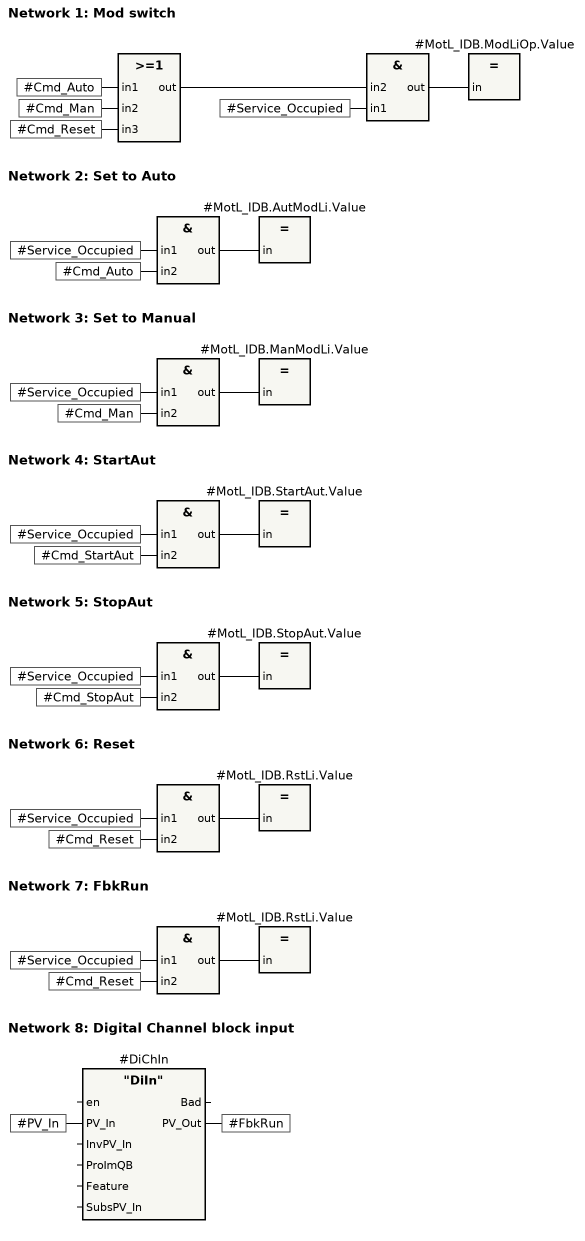
   #MotL_IDB.ModLiOp.Value := (#Cmd_Auto OR #Cmd_Man OR #Cmd_Reset) AND #Service_Occupied;
END_REGION

REGION Network 2: Set to Auto
   #MotL_IDB.AutModLi.Value := #Service_Occupied AND #Cmd_Auto;
END_REGION

REGION Network 3: Set to Manual
   #MotL_IDB.ManModLi.Value := #Service_Occupied AND #Cmd_Man;
END_REGION

REGION Network 4: StartAut
   #MotL_IDB.StartAut.Value := #Service_Occupied AND #Cmd_StartAut;
END_REGION

REGION Network 5: StopAut
   #MotL_IDB.StopAut.Value := #Service_Occupied AND #Cmd_StopAut;
END_REGION

REGION Network 6: Reset
   #MotL_IDB.RstLi.Value := #Service_Occupied AND #Cmd_Reset;
END_REGION

REGION Network 7: FbkRun
   #MotL_IDB.RstLi.Value := #Service_Occupied AND #Cmd_Reset;
END_REGION

REGION Network 8: Digital Channel block input
   #DiChIn(PV_In := #PV_In, PV_Out => #FbkRun);   // "DiIn"
END_REGION

REGION Network 9: CSF
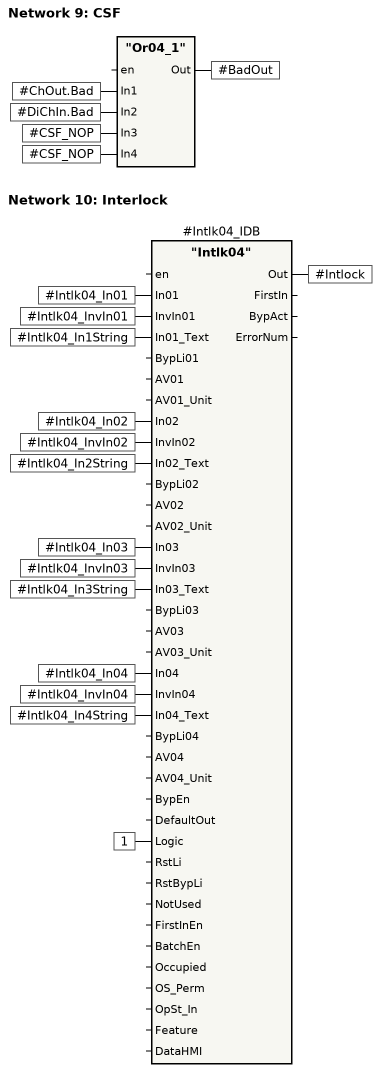
   "Or04_1"(In1 := #ChOut.Bad, In2 := #DiChIn.Bad, In3 := #CSF_NOP, In4 := #CSF_NOP, Out => #BadOut);
END_REGION

REGION Network 10: Interlock
   #Intlk04_IDB(In01 := #Intlk04_In01,   // "Intlk04"
                InvIn01 := #Intlk04_InvIn01,
                In01_Text := #Intlk04_In1String,
                In02 := #Intlk04_In02,
                InvIn02 := #Intlk04_InvIn02,
                In02_Text := #Intlk04_In2String,
                In03 := #Intlk04_In03,
                InvIn03 := #Intlk04_InvIn03,
                In03_Text := #Intlk04_In3String,
                In04 := #Intlk04_In04,
                InvIn04 := #Intlk04_InvIn04,
                In04_Text := #Intlk04_In4String,
                Logic := 1,
                Out => #Intlock);
END_REGION

REGION Network 11: MotSpdCL
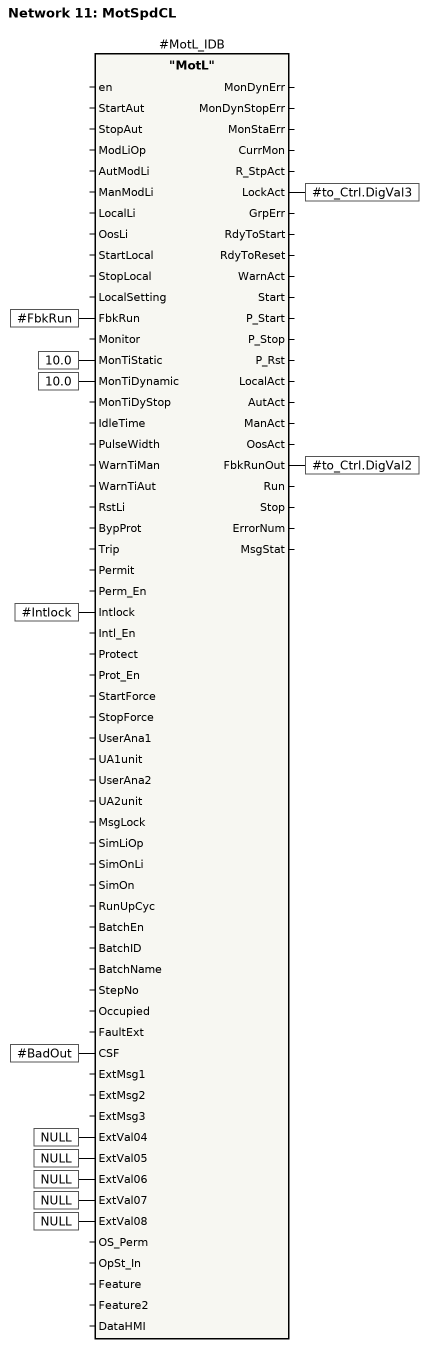
   #MotL_IDB(FbkRun := #FbkRun,   // "MotL"
             MonTiStatic := 10.0,
             MonTiDynamic := 10.0,
             Intlock := #Intlock,
             CSF := #BadOut,
             ExtVal04 := NULL,
             ExtVal05 := NULL,
             ExtVal06 := NULL,
             ExtVal07 := NULL,
             ExtVal08 := NULL,
             LockAct => #to_Ctrl.DigVal3,
             FbkRunOut => #to_Ctrl.DigVal2);
END_REGION

REGION Network 12: Channel block output
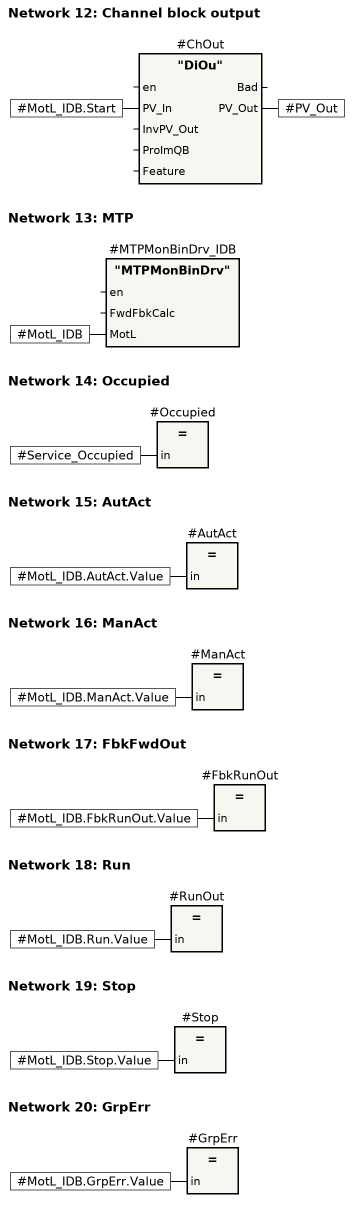
   #ChOut(PV_In := #MotL_IDB.Start, PV_Out => #PV_Out);   // "DiOu"
END_REGION

REGION Network 13: MTP
   #MTPMonBinDrv_IDB(MotL := #MotL_IDB);   // "MTPMonBinDrv"
END_REGION

REGION Network 14: Occupied
   #Occupied := #Service_Occupied;
END_REGION

REGION Network 15: AutAct
   #AutAct := #MotL_IDB.AutAct.Value;
END_REGION

REGION Network 16: ManAct
   #ManAct := #MotL_IDB.ManAct.Value;
END_REGION

REGION Network 17: FbkFwdOut
   #FbkRunOut := #MotL_IDB.FbkRunOut.Value;
END_REGION

REGION Network 18: Run
   #RunOut := #MotL_IDB.Run.Value;
END_REGION

REGION Network 19: Stop
   #Stop := #MotL_IDB.Stop.Value;
END_REGION

REGION Network 20: GrpErr
   #GrpErr := #MotL_IDB.GrpErr.Value;
END_REGION
END_FUNCTION_BLOCK

FUNCTION "P101" : Void   // FC17, FBD
{ S7_Optimized_Access := 'TRUE' }
// stored: SetENOAutomatically false
   VAR_TEMP
      Temp : "DigVal";
      Temp_1 : "DigVal";
      Temp_3 : "DigVal";
      Temp_2 : "DigVal";
      Temp_Error : "DigVal";
      In03 : "DigVal";
      State : "Service_States";
      FbkRun : "DigVal";
      StopAut : Bool;
   END_VAR
   VAR_TEMP   // added for the SCL form of the ladder/FBD networks
      _w1 : Bool;
   END_VAR
BEGIN

REGION Network 1: simulate Fbk Error
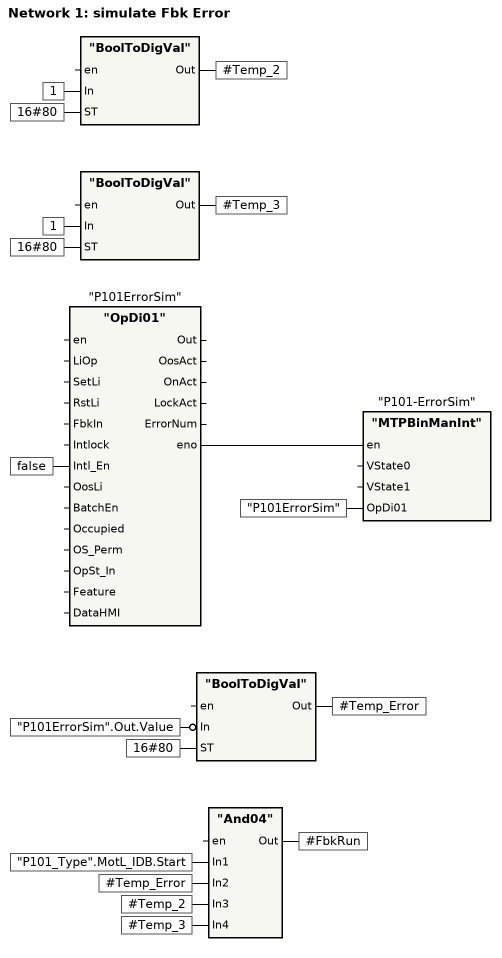
   "BoolToDigVal"(In := 1, ST := 16#80, Out => #Temp_2);
   "BoolToDigVal"(In := 1, ST := 16#80, Out => #Temp_3);
   "P101ErrorSim"(Intl_En := false, ENO => #_w1);   // "OpDi01"
   IF #_w1 THEN
       "P101-ErrorSim"(OpDi01 := "P101ErrorSim");   // "MTPBinManInt"
   END_IF;
   "BoolToDigVal"(In := NOT "P101ErrorSim".Out.Value, ST := 16#80, Out => #Temp_Error);
   "And04"(In1 := "P101_Type".MotL_IDB.Start,
           In2 := #Temp_Error,
           In3 := #Temp_2,
           In4 := #Temp_3,
           Out => #FbkRun);
END_REGION

REGION Network 2: Pump interconnections
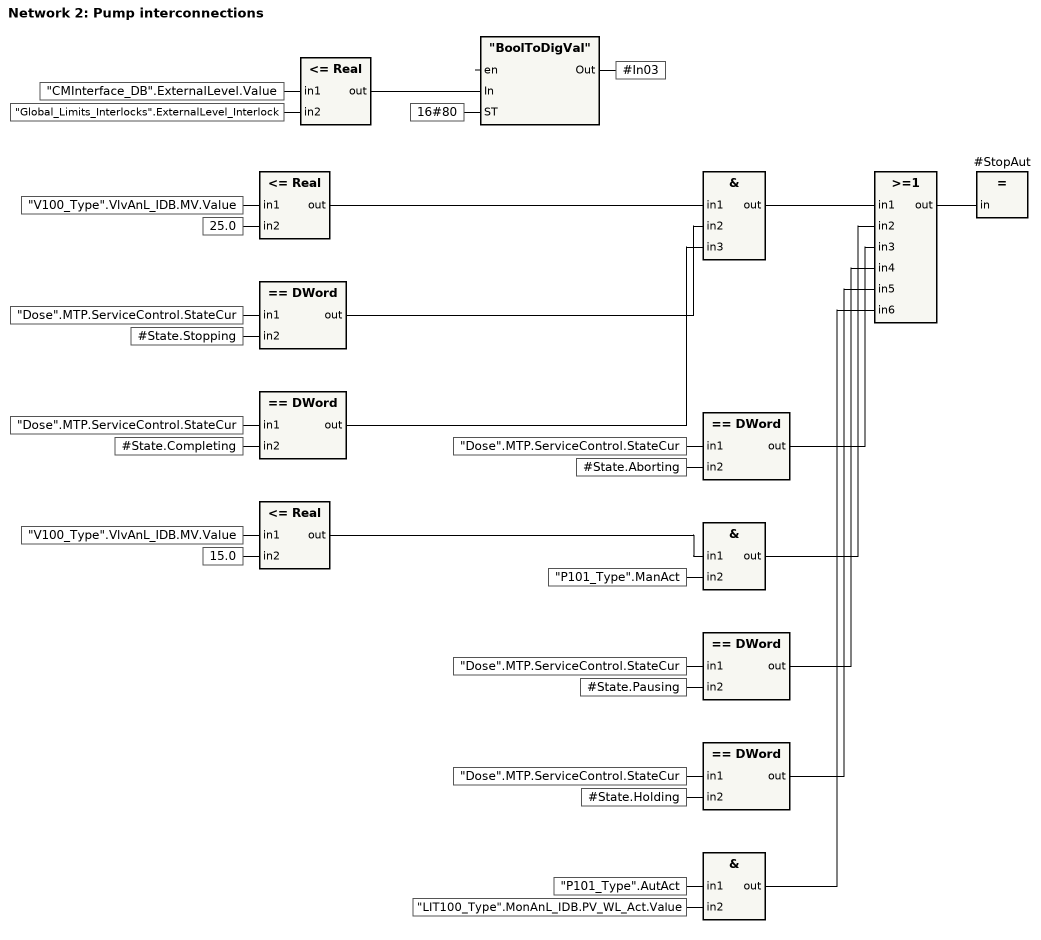
   "BoolToDigVal"(In := "CMInterface_DB".ExternalLevel.Value <= "Global_Limits_Interlocks".ExternalLevel_Interlock,
                  ST := 16#80,
                  Out => #In03);
   #StopAut := (("V100_Type".VlvAnL_IDB.MV.Value <= 25.0) AND ("Dose".MTP.ServiceControl.StateCur = #State.Stopping) AND ("Dose".MTP.ServiceControl.StateCur = #State.Completing)) OR (("V100_Type".VlvAnL_IDB.MV.Value <= 15.0) AND "P101_Type".ManAct) OR ("Dose".MTP.ServiceControl.StateCur = #State.Aborting) OR ("Dose".MTP.ServiceControl.StateCur = #State.Pausing) OR ("Dose".MTP.ServiceControl.StateCur = #State.Holding) OR ("P101_Type".AutAct AND "LIT100_Type".MonAnL_IDB.PV_WL_Act.Value);
END_REGION

REGION Network 3: MotL
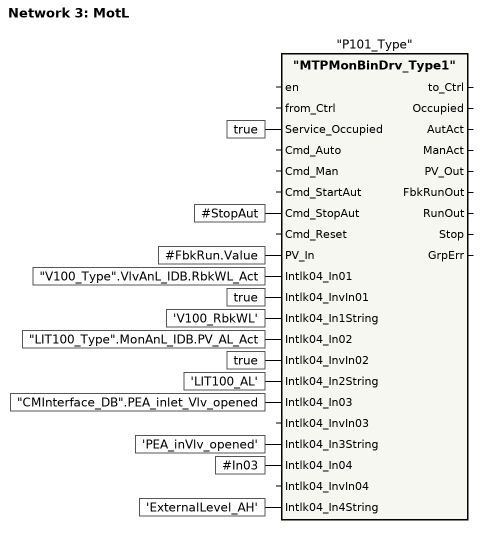
   "P101_Type"(Service_Occupied := true,   // "MTPMonBinDrv_Type1"
               Cmd_StopAut := #StopAut,
               PV_In := #FbkRun.Value,
               Intlk04_In01 := "V100_Type".VlvAnL_IDB.RbkWL_Act,
               Intlk04_InvIn01 := true,
               Intlk04_In1String := 'V100_RbkWL',
               Intlk04_In02 := "LIT100_Type".MonAnL_IDB.PV_AL_Act,
               Intlk04_InvIn02 := true,
               Intlk04_In2String := 'LIT100_AL',
               Intlk04_In03 := "CMInterface_DB".PEA_inlet_Vlv_opened,
               Intlk04_In3String := 'PEA_inVlv_opened',
               Intlk04_In04 := #In03,
               Intlk04_In4String := 'ExternalLevel_AH');
END_REGION
END_FUNCTION

FUNCTION "V100" : Void   // FC3, FBD
{ S7_Optimized_Access := 'TRUE' }
// stored: SetENOAutomatically false
   VAR_TEMP
      Temp : "DigVal";
      In03 : "DigVal";
      Temp_FF : "DigVal";
      Temp_fromCTRL : "StruCm";
   END_VAR
BEGIN

REGION Network 1: VlvAnL interconnections
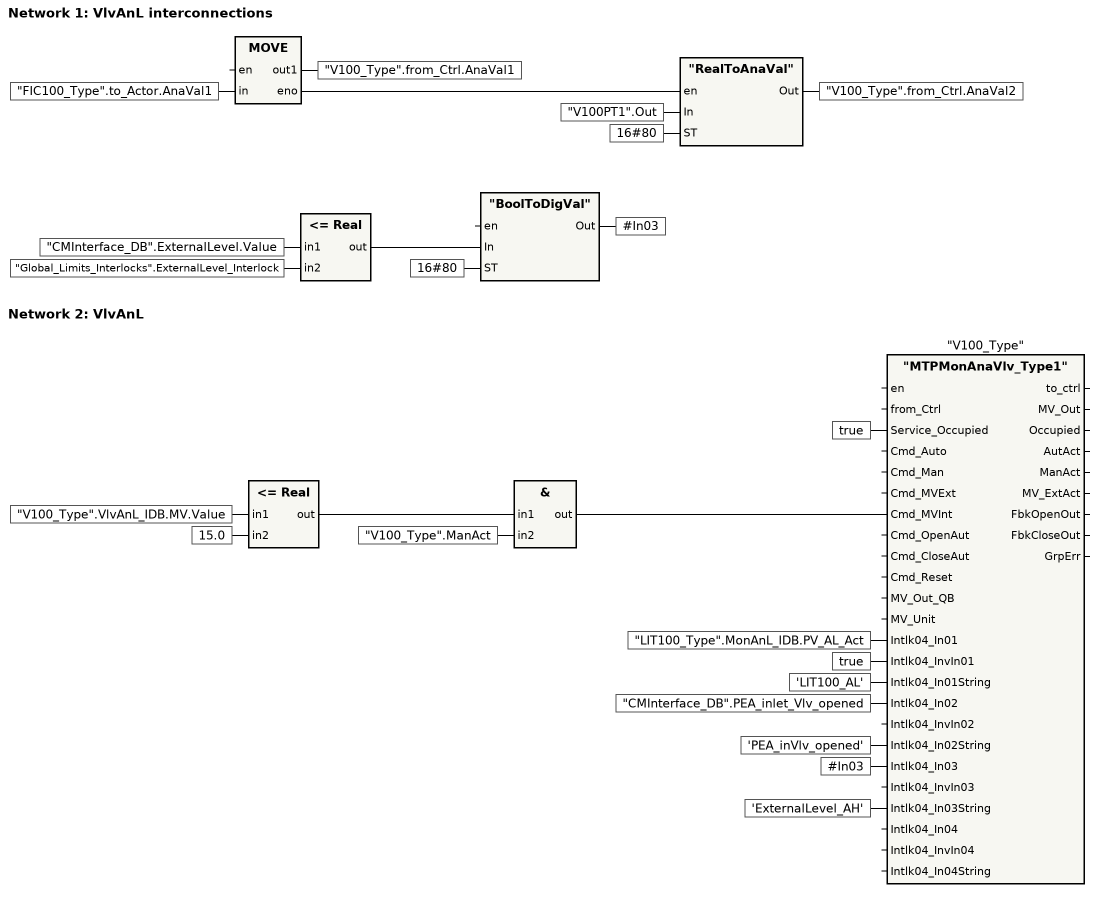
   "V100_Type".from_Ctrl.AnaVal1 := "FIC100_Type".to_Actor.AnaVal1;
   "RealToAnaVal"(In := "V100PT1".Out, ST := 16#80, Out => "V100_Type".from_Ctrl.AnaVal2);
   "BoolToDigVal"(In := "CMInterface_DB".ExternalLevel.Value <= "Global_Limits_Interlocks".ExternalLevel_Interlock,
                  ST := 16#80,
                  Out => #In03);
END_REGION

REGION Network 2: VlvAnL
   "V100_Type"(Service_Occupied := true,   // "MTPMonAnaVlv_Type1"
               Cmd_MVInt := ("V100_Type".VlvAnL_IDB.MV.Value <= 15.0) AND "V100_Type".ManAct,
               Intlk04_In01 := "LIT100_Type".MonAnL_IDB.PV_AL_Act,
               Intlk04_InvIn01 := true,
               Intlk04_In01String := 'LIT100_AL',
               Intlk04_In02 := "CMInterface_DB".PEA_inlet_Vlv_opened,
               Intlk04_In02String := 'PEA_inVlv_opened',
               Intlk04_In03 := #In03,
               Intlk04_In03String := 'ExternalLevel_AH');
END_REGION
END_FUNCTION

FUNCTION "RealToAnaVal" : Void   // FC9, SCL
{ S7_Optimized_Access := 'TRUE' }
// stored: SetENOAutomatically false
   VAR_INPUT
      In : Real;
      ST : Byte;
   END_VAR
   VAR_OUTPUT
      Out : "AnaVal";
   END_VAR
BEGIN
   #Out.ST := #ST;
   #Out.Value := #In;
END_FUNCTION

FUNCTION_BLOCK "MTPMonAnaVlv_Type1"   // FB7, FBD
{ S7_Optimized_Access := 'TRUE' }
// stored: MemoryReserve 100, SetENOAutomatically false
   VAR_INPUT
      from_Ctrl { ExternalAccessible := 'False'; ExternalVisible := 'False'; ExternalWritable := 'False'} : "StruCm";
      Service_Occupied { ExternalAccessible := 'False'; ExternalVisible := 'False'; ExternalWritable := 'False'} : Bool;
      Cmd_Auto { ExternalAccessible := 'False'; ExternalVisible := 'False'; ExternalWritable := 'False'} : Bool;
      Cmd_Man { ExternalAccessible := 'False'; ExternalVisible := 'False'; ExternalWritable := 'False'} : Bool;
      Cmd_MVExt { ExternalAccessible := 'False'; ExternalVisible := 'False'; ExternalWritable := 'False'} : Bool;
      Cmd_MVInt { ExternalAccessible := 'False'; ExternalVisible := 'False'; ExternalWritable := 'False'} : Bool;
      Cmd_OpenAut { ExternalAccessible := 'False'; ExternalVisible := 'False'; ExternalWritable := 'False'} : Bool;
      Cmd_CloseAut { ExternalAccessible := 'False'; ExternalVisible := 'False'; ExternalWritable := 'False'} : Bool;
      Cmd_Reset { ExternalAccessible := 'False'; ExternalVisible := 'False'; ExternalWritable := 'False'} : Bool;
      MV_Out_QB { ExternalAccessible := 'False'; ExternalVisible := 'False'; ExternalWritable := 'False'} : Bool := true;
      MV_Unit { ExternalAccessible := 'False'; ExternalVisible := 'False'; ExternalWritable := 'False'} : Int := 1342;
      Intlk04_In01 { ExternalAccessible := 'False'; ExternalVisible := 'False'; ExternalWritable := 'False'} : "DigVal";
      Intlk04_InvIn01 { ExternalAccessible := 'False'; ExternalVisible := 'False'; ExternalWritable := 'False'} : Bool;
      Intlk04_In01String : String;
      Intlk04_In02 { ExternalAccessible := 'False'; ExternalVisible := 'False'; ExternalWritable := 'False'} : "DigVal";
      Intlk04_InvIn02 { ExternalAccessible := 'False'; ExternalVisible := 'False'; ExternalWritable := 'False'} : Bool;
      Intlk04_In02String : String;
      Intlk04_In03 { ExternalAccessible := 'False'; ExternalVisible := 'False'; ExternalWritable := 'False'} : "DigVal";
      Intlk04_InvIn03 { ExternalAccessible := 'False'; ExternalVisible := 'False'; ExternalWritable := 'False'} : Bool;
      Intlk04_In03String : String;
      Intlk04_In04 { ExternalAccessible := 'False'; ExternalVisible := 'False'; ExternalWritable := 'False'} : "DigVal";
      Intlk04_InvIn04 { ExternalAccessible := 'False'; ExternalVisible := 'False'; ExternalWritable := 'False'} : Bool;
      Intlk04_In04String : String;
   END_VAR
   VAR_OUTPUT
      to_ctrl { ExternalAccessible := 'False'; ExternalVisible := 'False'; ExternalWritable := 'False'} : "StruCm";
      MV_Out { ExternalAccessible := 'False'; ExternalVisible := 'False'; ExternalWritable := 'False'} : Word;
      Occupied { ExternalAccessible := 'False'; ExternalVisible := 'False'; ExternalWritable := 'False'} : Bool;   // Occupied by a Service procedure
      AutAct { ExternalAccessible := 'False'; ExternalVisible := 'False'; ExternalWritable := 'False'} : Bool;
      ManAct { ExternalAccessible := 'False'; ExternalVisible := 'False'; ExternalWritable := 'False'} : Bool;
      MV_ExtAct { ExternalAccessible := 'False'; ExternalVisible := 'False'; ExternalWritable := 'False'} : Bool;
      FbkOpenOut { ExternalAccessible := 'False'; ExternalVisible := 'False'; ExternalWritable := 'False'} : Bool;
      FbkCloseOut { ExternalAccessible := 'False'; ExternalVisible := 'False'; ExternalWritable := 'False'} : Bool;
      GrpErr { ExternalAccessible := 'False'; ExternalVisible := 'False'; ExternalWritable := 'False'} : Bool;
   END_VAR
   VAR
      AnOut_IDB { ExternalAccessible := 'False'; ExternalVisible := 'False'; ExternalWritable := 'False'} : "AnOu";
      Intlk04_IDB : "Intlk04";
      VlvAnL_IDB { S7_SetPoint := 'True'} : "VlvAnL";
      MTPMonAnaVlv_IDB { ExternalVisible := 'False'; S7_SetPoint := 'True'} : "MTPMonAnaVlv";
   END_VAR
   VAR_TEMP
      CSF_NOP : "DigVal";
      BadAnIn : "DigVal";
      BadOut : "DigVal";
      Intlock : "DigVal";
   END_VAR
   // Intlk04_In01.Value := true;
   // Intlk04_In02.Value := true;
   // Intlk04_In03.Value := true;
   // Intlk04_In04.Value := true;
BEGIN

REGION Network 1: Convert
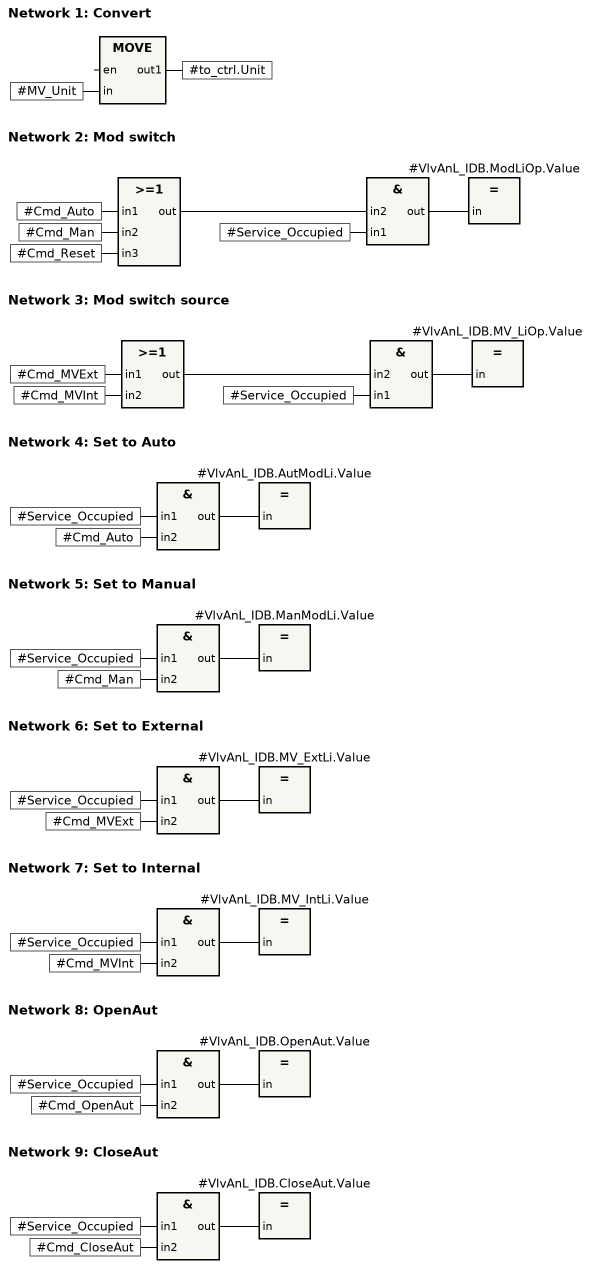
   #to_ctrl.Unit := #MV_Unit;
END_REGION

REGION Network 2: Mod switch
   #VlvAnL_IDB.ModLiOp.Value := (#Cmd_Auto OR #Cmd_Man OR #Cmd_Reset) AND #Service_Occupied;
END_REGION

REGION Network 3: Mod switch source
   #VlvAnL_IDB.MV_LiOp.Value := (#Cmd_MVExt OR #Cmd_MVInt) AND #Service_Occupied;
END_REGION

REGION Network 4: Set to Auto
   #VlvAnL_IDB.AutModLi.Value := #Service_Occupied AND #Cmd_Auto;
END_REGION

REGION Network 5: Set to Manual
   #VlvAnL_IDB.ManModLi.Value := #Service_Occupied AND #Cmd_Man;
END_REGION

REGION Network 6: Set to External
   #VlvAnL_IDB.MV_ExtLi.Value := #Service_Occupied AND #Cmd_MVExt;
END_REGION

REGION Network 7: Set to Internal
   #VlvAnL_IDB.MV_IntLi.Value := #Service_Occupied AND #Cmd_MVInt;
END_REGION

REGION Network 8: OpenAut
   #VlvAnL_IDB.OpenAut.Value := #Service_Occupied AND #Cmd_OpenAut;
END_REGION

REGION Network 9: CloseAut
   #VlvAnL_IDB.CloseAut.Value := #Service_Occupied AND #Cmd_CloseAut;
END_REGION

REGION Network 10: Reset
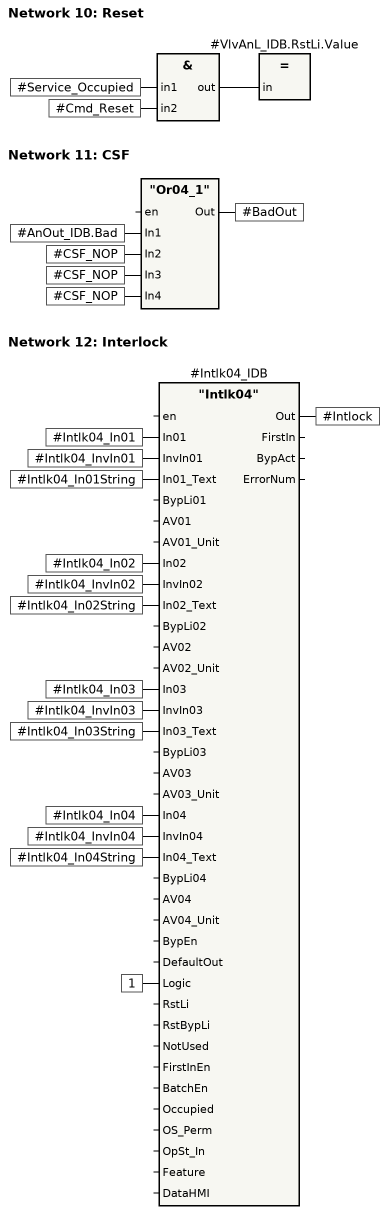
   #VlvAnL_IDB.RstLi.Value := #Service_Occupied AND #Cmd_Reset;
END_REGION

REGION Network 11: CSF
   "Or04_1"(In1 := #AnOut_IDB.Bad, In2 := #CSF_NOP, In3 := #CSF_NOP, In4 := #CSF_NOP, Out => #BadOut);
END_REGION

REGION Network 12: Interlock
   #Intlk04_IDB(In01 := #Intlk04_In01,   // "Intlk04"
                InvIn01 := #Intlk04_InvIn01,
                In01_Text := #Intlk04_In01String,
                In02 := #Intlk04_In02,
                InvIn02 := #Intlk04_InvIn02,
                In02_Text := #Intlk04_In02String,
                In03 := #Intlk04_In03,
                InvIn03 := #Intlk04_InvIn03,
                In03_Text := #Intlk04_In03String,
                In04 := #Intlk04_In04,
                InvIn04 := #Intlk04_InvIn04,
                In04_Text := #Intlk04_In04String,
                Logic := 1,
                Out => #Intlock);
END_REGION

REGION Network 13: VlvAnL
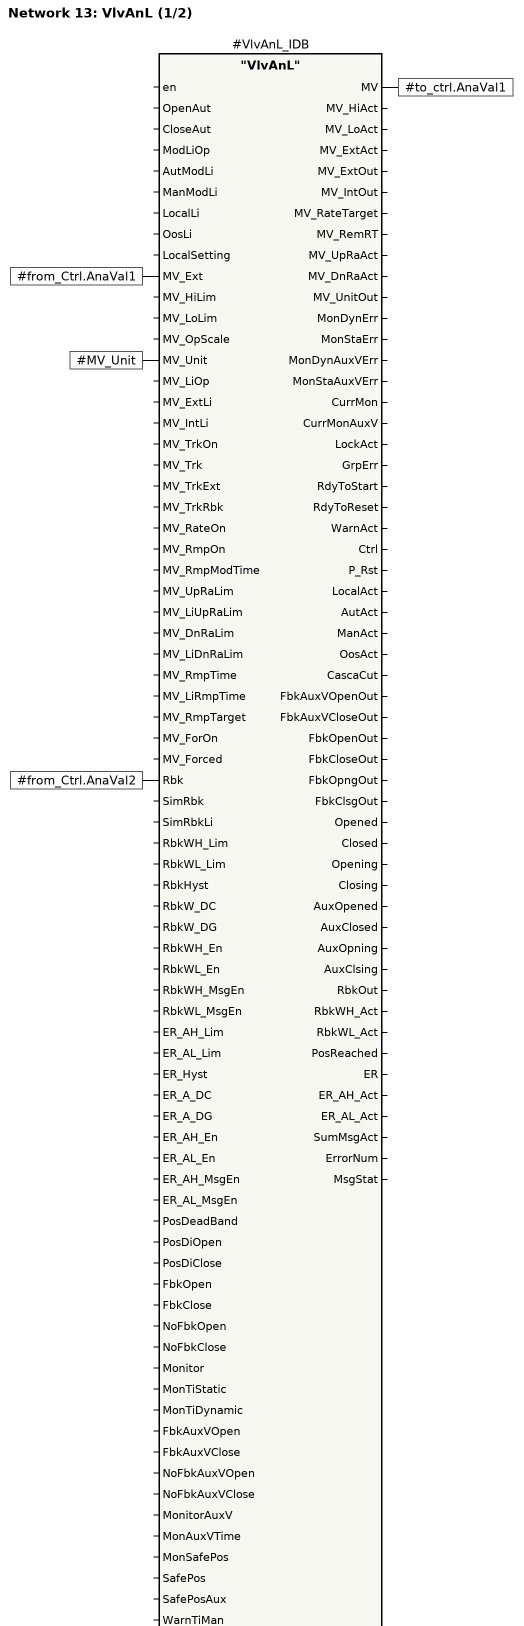
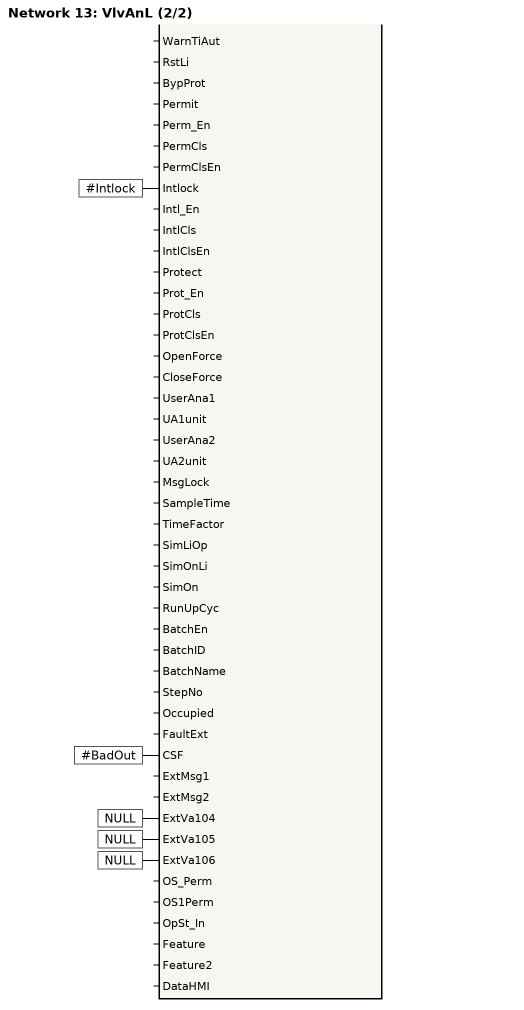
   #VlvAnL_IDB(MV_Ext := #from_Ctrl.AnaVal1,   // "VlvAnL"
               MV_Unit := #MV_Unit,
               Rbk := #from_Ctrl.AnaVal2,
               Intlock := #Intlock,
               CSF := #BadOut,
               ExtVa104 := NULL,
               ExtVa105 := NULL,
               ExtVa106 := NULL,
               MV => #to_ctrl.AnaVal1);
END_REGION

REGION Network 14: Analog Out
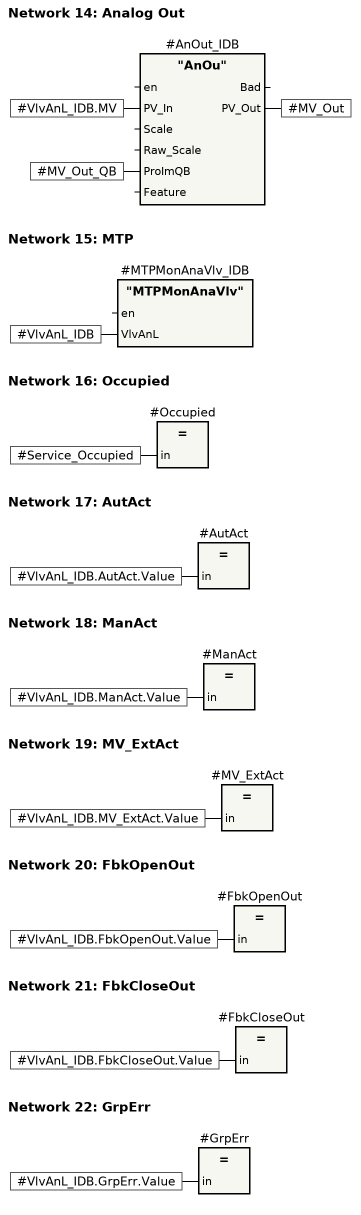
   #AnOut_IDB(PV_In := #VlvAnL_IDB.MV, ProImQB := #MV_Out_QB, PV_Out => #MV_Out);   // "AnOu"
END_REGION

REGION Network 15: MTP
   #MTPMonAnaVlv_IDB(VlvAnL := #VlvAnL_IDB);   // "MTPMonAnaVlv"
END_REGION

REGION Network 16: Occupied
   #Occupied := #Service_Occupied;
END_REGION

REGION Network 17: AutAct
   #AutAct := #VlvAnL_IDB.AutAct.Value;
END_REGION

REGION Network 18: ManAct
   #ManAct := #VlvAnL_IDB.ManAct.Value;
END_REGION

REGION Network 19: MV_ExtAct
   #MV_ExtAct := #VlvAnL_IDB.MV_ExtAct.Value;
END_REGION

REGION Network 20: FbkOpenOut
   #FbkOpenOut := #VlvAnL_IDB.FbkOpenOut.Value;
END_REGION

REGION Network 21: FbkCloseOut
   #FbkCloseOut := #VlvAnL_IDB.FbkCloseOut.Value;
END_REGION

REGION Network 22: GrpErr
   #GrpErr := #VlvAnL_IDB.GrpErr.Value;
END_REGION
END_FUNCTION_BLOCK

FUNCTION "Flow_Sim" : Void   // FC14, FBD
{ S7_Optimized_Access := 'TRUE' }
// stored: SetENOAutomatically false
   VAR_TEMP
      State : "Service_States";
   END_VAR
BEGIN

REGION Network 1: flow value
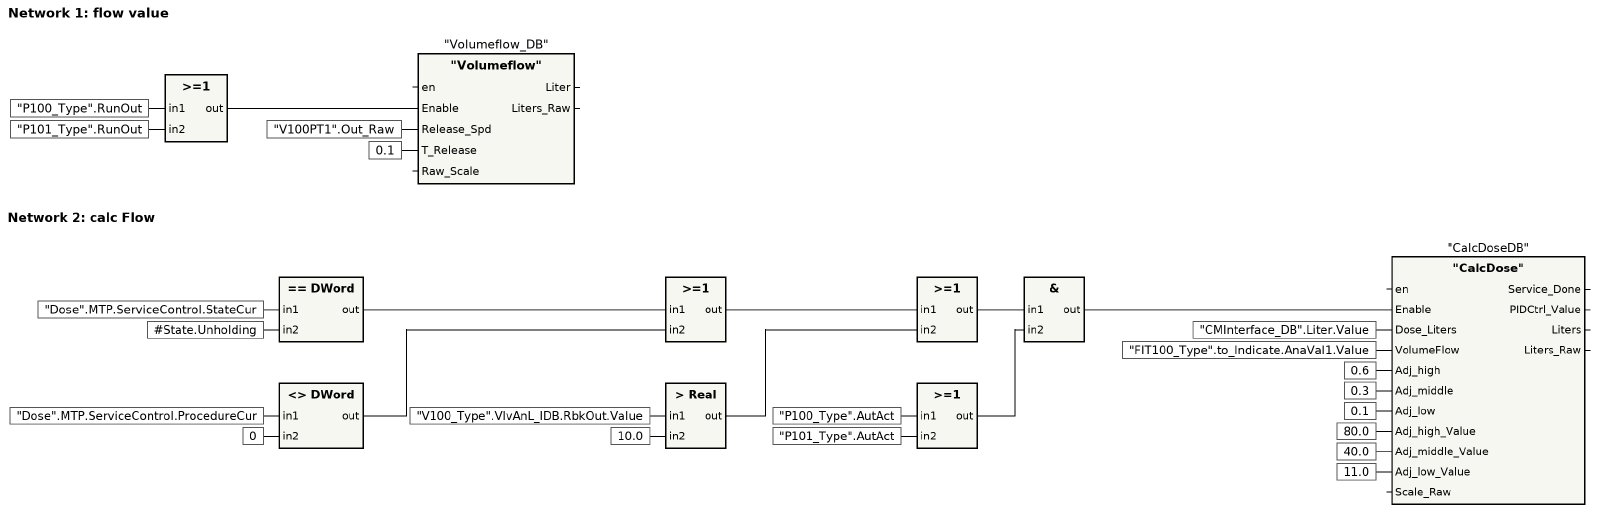
   "Volumeflow_DB"(Enable := "P100_Type".RunOut OR "P101_Type".RunOut,   // "Volumeflow"
                   Release_Spd := "V100PT1".Out_Raw,
                   T_Release := 0.1);
END_REGION

REGION Network 2: calc Flow
   "CalcDoseDB"(Enable := (("Dose".MTP.ServiceControl.StateCur = #State.Unholding) OR ("Dose".MTP.ServiceControl.ProcedureCur <> 0) OR ("V100_Type".VlvAnL_IDB.RbkOut.Value > 10.0)) AND ("P100_Type".AutAct OR "P101_Type".AutAct),   // "CalcDose"
                Dose_Liters := "CMInterface_DB".Liter.Value,
                VolumeFlow := "FIT100_Type".to_Indicate.AnaVal1.Value,
                Adj_high := 0.6,
                Adj_middle := 0.3,
                Adj_low := 0.1,
                Adj_high_Value := 80.0,
                Adj_middle_Value := 40.0,
                Adj_low_Value := 11.0);
END_REGION
END_FUNCTION

FUNCTION_BLOCK "Volumeflow"   // FB1, SCL
{ S7_Optimized_Access := 'TRUE' }
// stored: MemoryReserve 100, SetENOAutomatically false
   VAR_INPUT
      Enable : Bool;
      Release_Spd : Int;
      T_Release : Real;
      Raw_Scale { ExternalAccessible := 'False'; ExternalVisible := 'False'; ExternalWritable := 'False'} : "ScaVal_Raw";
   END_VAR
   VAR_OUTPUT
      Liter : Real;
      Liters_Raw : Int;
   END_VAR
   VAR
      pi : Real := 3.1415;
      r : Real := 0.5;
   END_VAR
   VAR_TEMP
      Release_Spd_Raw : Real;
      Release_Spd_Real : Real;
   END_VAR
   // Raw_Scale.High := 27648;
   // Raw_Scale.Low := 0;
BEGIN
   IF #Enable = FALSE THEN
       #Liter := 0;
       #Liters_Raw := 0;
       RETURN;
   END_IF;
   #Release_Spd_Real := INT_TO_REAL(#Release_Spd);
   #Release_Spd_Raw := (#Release_Spd_Real / 27648) * 100;
   //Volume flow in liter (dm^2 == l)
   #Liter := #T_Release * #Release_Spd_Raw * #pi * #r * #r * 4;
   #Liters_Raw := (#Liter/32) * #Raw_Scale.High;
END_FUNCTION_BLOCK

FUNCTION_BLOCK "CalcDose"   // FB2, SCL
{ S7_Optimized_Access := 'TRUE' }
// stored: MemoryReserve 100, SetENOAutomatically false
   VAR_INPUT
      Enable : Bool;
      Dose_Liters : Real;
      VolumeFlow : Real;
      Adj_high : Real;
      Adj_middle : Real;
      Adj_low : Real;
      Adj_high_Value : Real;
      Adj_middle_Value : Real;
      Adj_low_Value : Real;
      Scale_Raw : "ScaVal_Raw";
   END_VAR
   VAR_OUTPUT
      Service_Done : Bool;
      PIDCtrl_Value : "AnaVal";
      Liters { ExternalWritable := 'False'} : Real;
      Liters_Raw : Int;
   END_VAR
   VAR_TEMP
      Liters_Diff : Real;
      State : "Service_States";
   END_VAR
   // Scale_Raw.High := 27648;
   // Scale_Raw.Low := 0;
BEGIN
   IF "Dose".Information.state = #State.Starting THEN
       #Liters := 0;
       "AccuSDB".RstCnt1Li.ST := 16#80;
       "AccuSDB".RstCnt1Li.Value := TRUE;
       #Service_Done := FALSE;
   ELSE
       "AccuSDB".RstCnt1Li.ST := 16#80;
       "AccuSDB".RstCnt1Li.Value := False;
   END_IF;
   IF #Enable = FALSE THEN
       RETURN;
   END_IF;

   #PIDCtrl_Value.ST := 16#80;
   "AccuSDB".RstCnt1Li.ST := 16#80;
   //calc already pumped liters and set valve MV
   IF "Dose".Information.state = #State.Execute THEN
       //set valve MV for Procedure doseToEmpty
       IF "Dose".MTP.ServiceControl.ProcedureCur = 3 THEN
           "AccuSDB".RstCnt1Li.Value := False;
           #Liters := "AccuSDB".AcCnt1Out.Value;
           #PIDCtrl_Value.Value := 100;
           #Liters_Diff := #Dose_Liters - #Liters;
           IF "LIT100_Type".to_Indicate.AnaVal1.Value <= 1.0 THEN
               #PIDCtrl_Value.Value := 60;
           ELSIF "LIT100_Type".to_Indicate.AnaVal1.Value <= 0.5 THEN
               #PIDCtrl_Value.Value := 0;
           END_IF;
       //set valve MV for Procedure doseByFlow and DoseByVolume
       ELSE
           IF #Liters <= #Dose_Liters THEN
               #Liters := "AccuSDB".AcCnt1Out.Value;
           ELSIF #Liters > #Dose_Liters THEN
               #Service_Done := TRUE;
           END_IF;

           //calc PID ctrl value. Different MV depending on already pumped liters. 
           #Liters_Diff := #Dose_Liters - #Liters;
           IF "LIT100_Type".to_Indicate.AnaVal1.Value <= 0.4 OR #Liters_Diff = 0 THEN
               #PIDCtrl_Value.Value := 0;
           ELSIF #Liters_Diff <= #Adj_low * #Dose_Liters THEN
               #PIDCtrl_Value.Value := #Adj_low_Value;
           ELSIF #Liters_Diff <= (#Adj_middle * #Dose_Liters) AND #Liters_Diff > (#Adj_low * #Dose_Liters) THEN
               #PIDCtrl_Value.Value := #Adj_middle_Value;
           ELSIF #Liters_Diff <= (#Adj_high * #Dose_Liters) AND #Liters_Diff > (#Adj_middle * #Dose_Liters) THEN
               #PIDCtrl_Value.Value := #Adj_high_Value;
           ELSE
               #PIDCtrl_Value.Value := 100;
           END_IF;
       END_IF;
   ELSIF "Dose".Information.state <> #State.Execute THEN
       #PIDCtrl_Value.Value := 0;
   END_IF;

   #Liters_Raw := (#Liters/3600) * #Scale_Raw.High;
END_FUNCTION_BLOCK

FUNCTION "Level_Sim" : Void   // FC1, FBD
{ S7_Optimized_Access := 'TRUE' }
// stored: SetENOAutomatically false
   VAR_TEMP   // added for the SCL form of the ladder/FBD networks
      _w1 : Bool;
   END_VAR
BEGIN

REGION Network 1: LevelSimulation
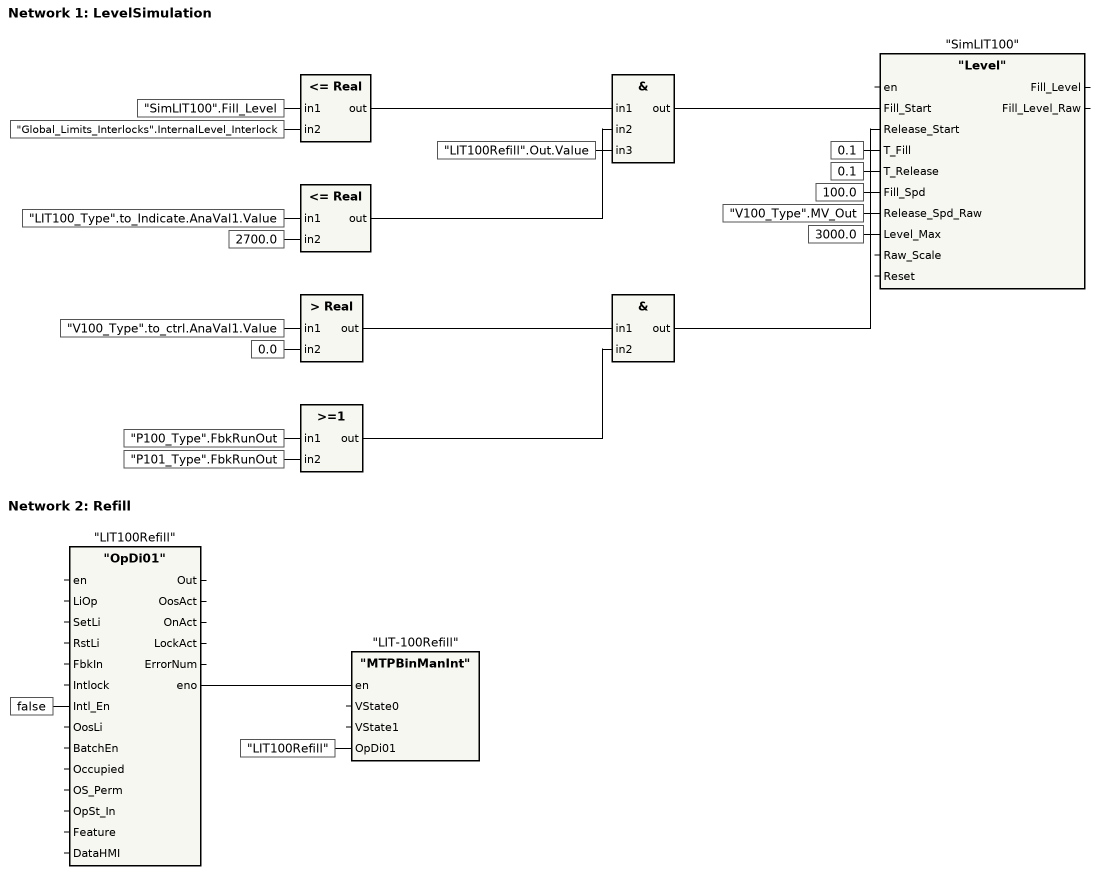
   "SimLIT100"(Fill_Start := ("SimLIT100".Fill_Level <= "Global_Limits_Interlocks".InternalLevel_Interlock) AND ("LIT100_Type".to_Indicate.AnaVal1.Value <= 2700.0) AND "LIT100Refill".Out.Value,   // "Level"
               Release_Start := ("V100_Type".to_ctrl.AnaVal1.Value > 0.0) AND ("P100_Type".FbkRunOut OR "P101_Type".FbkRunOut),
               T_Fill := 0.1,
               T_Release := 0.1,
               Fill_Spd := 100.0,
               Release_Spd_Raw := "V100_Type".MV_Out,
               Level_Max := 3000.0);
END_REGION

REGION Network 2: Refill
   "LIT100Refill"(Intl_En := false, ENO => #_w1);   // "OpDi01"
   IF #_w1 THEN
       "LIT-100Refill"(OpDi01 := "LIT100Refill");   // "MTPBinManInt"
   END_IF;
END_REGION
END_FUNCTION

FUNCTION_BLOCK "Level"   // FB11, SCL
{ S7_Optimized_Access := 'TRUE' }
// stored: MemoryReserve 100, SetENOAutomatically false
   VAR_INPUT
      Fill_Start { ExternalAccessible := 'False'; ExternalVisible := 'False'; ExternalWritable := 'False'} : Bool;   // 1 = Starts fill process
      Release_Start { ExternalAccessible := 'False'; ExternalVisible := 'False'; ExternalWritable := 'False'} : Bool;   // 1 = Starts release prozess
      T_Fill { ExternalAccessible := 'False'; ExternalVisible := 'False'; ExternalWritable := 'False'} : Real := 1.0;   // Time constant
      T_Release { ExternalAccessible := 'False'; ExternalVisible := 'False'; ExternalWritable := 'False'} : Real := 1.0;   // Execution cycle @ OB3x. E.g. 100 ms = 0.1s
      Fill_Spd { ExternalAccessible := 'False'; ExternalVisible := 'False'; ExternalWritable := 'False'} : Real := 100.0;   // Filling speed in %
      Release_Spd_Raw { ExternalAccessible := 'False'; ExternalVisible := 'False'; ExternalWritable := 'False'} : Int := 27648;   // Releasing speed in %
      Level_Max { ExternalAccessible := 'False'; ExternalVisible := 'False'; ExternalWritable := 'False'} : Real := 100.0;   // Max Level
      Raw_Scale { ExternalAccessible := 'False'; ExternalVisible := 'False'; ExternalWritable := 'False'} : "ScaVal_Raw";
      Reset { ExternalAccessible := 'False'; ExternalVisible := 'False'; ExternalWritable := 'False'} : Bool := False;   // Reset level to 0.0
   END_VAR
   VAR_OUTPUT
      Fill_Level { ExternalAccessible := 'False'; ExternalVisible := 'False'; ExternalWritable := 'False'} : Real := 1500.0;
      Fill_Level_Raw { ExternalAccessible := 'False'; ExternalVisible := 'False'; ExternalWritable := 'False'} : Int;
   END_VAR
   VAR_TEMP
      Release_Spd : Real;
      ReleaseSpd_Real : Real;
   END_VAR
   // Raw_Scale.High := 27648;
   // Raw_Scale.Low := 0;
BEGIN
   #ReleaseSpd_Real := INT_TO_REAL(#Release_Spd_Raw);
   #Release_Spd := (#ReleaseSpd_Real / 27648) * 100;

   // Fill
   IF #Fill_Start = True AND #Fill_Level <= #Level_Max THEN
       #Fill_Level := #Fill_Level + (#T_Fill * (#Fill_Spd) * 3.1);
   END_IF;

   // Release
   IF #Release_Start = True AND #Fill_Level >= 0.0 THEN
       #Fill_Level := #Fill_Level - (#T_Release * (#Release_Spd / 10.0 * 3.1));
   END_IF;

   // Prevent negative fill level / Reset
   IF #Fill_Level < 0.0 OR #Reset = True THEN
       #Fill_Level := 0.0;
   END_IF;

   // Prevent overfilling
   IF #Fill_Level > #Level_Max THEN
       #Fill_Level := #Level_Max;
   END_IF;

   // Raw output
   #Fill_Level_Raw := ((#Fill_Level / #Level_Max) * #Raw_Scale.High);
END_FUNCTION_BLOCK

FUNCTION "Vlv_Sim" : Void   // FC13, FBD
{ S7_Optimized_Access := 'TRUE' }
// stored: SetENOAutomatically false
BEGIN

REGION Network 1: PT1
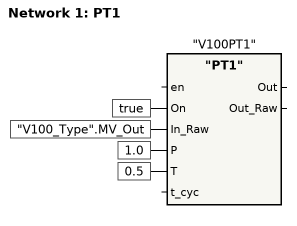
   "V100PT1"(On := true, In_Raw := "V100_Type".MV_Out, P := 1.0, T := 0.5);   // "PT1"
END_REGION
END_FUNCTION

FUNCTION_BLOCK "PT1"   // FB4, SCL
{ S7_Optimized_Access := 'TRUE' }
// stored: MemoryReserve 100, SetENOAutomatically false
   VAR_INPUT
      On { ExternalAccessible := 'False'; ExternalVisible := 'False'; ExternalWritable := 'False'} : Bool;   // 0 = Off => In = 0.0
      In_Raw { ExternalAccessible := 'False'; ExternalVisible := 'False'; ExternalWritable := 'False'} : Int;
      P { ExternalAccessible := 'False'; ExternalVisible := 'False'; ExternalWritable := 'False'} : Real := 1.0;   // Propotional parameter
      T { ExternalAccessible := 'False'; ExternalVisible := 'False'; ExternalWritable := 'False'} : Real := 1.0;   // Time constant [s]
      t_cyc { ExternalAccessible := 'False'; ExternalVisible := 'False'; ExternalWritable := 'False'} : Real := 0.1;   // OB-Cycle time
   END_VAR
   VAR_OUTPUT
      Out { ExternalAccessible := 'False'; ExternalVisible := 'False'; ExternalWritable := 'False'} : Real := 0.0;
      Out_Raw : Int := 0;
   END_VAR
   VAR
      "Out-1" { ExternalAccessible := 'False'; ExternalVisible := 'False'; ExternalWritable := 'False'} : Real := 0.0;
   END_VAR
BEGIN
   IF #On THEN
       #Out_Raw := #"Out-1" + (#P * (#In_Raw - #"Out-1") * (#t_cyc / (#T + #t_cyc)));
   ELSE
       #Out_Raw := #"Out-1" + (#P * (0.0 - #"Out-1") * (#t_cyc / (#T + #t_cyc)));
   END_IF;

   #"Out-1" := #Out_Raw; //Save output value end of this cycle
   #Out := (INT_TO_REAL(#Out_Raw) / 27648) * 100;
END_FUNCTION_BLOCK

FUNCTION "AccuS_Liter" : Void   // FC12, FBD
{ S7_Optimized_Access := 'TRUE' }
// stored: SetENOAutomatically false
   VAR_TEMP
      State : "Service_States";
   END_VAR
   VAR_TEMP   // added for the SCL form of the ladder/FBD networks
      _w1 : Bool;
   END_VAR
BEGIN

REGION Network 1
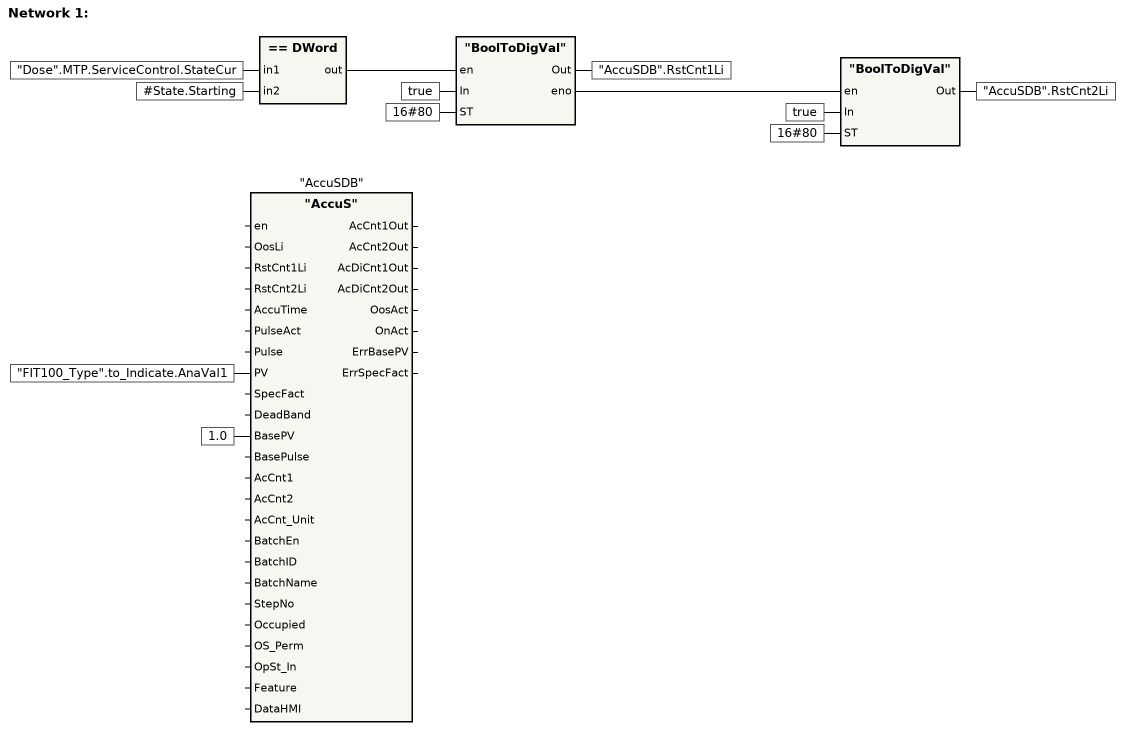
   "BoolToDigVal"(EN := "Dose".MTP.ServiceControl.StateCur = #State.Starting,
                  In := true,
                  ST := 16#80,
                  Out => "AccuSDB".RstCnt1Li,
                  ENO => #_w1);
   IF #_w1 THEN "BoolToDigVal"(In := true, ST := 16#80, Out => "AccuSDB".RstCnt2Li); END_IF;
   "AccuSDB"(PV := "FIT100_Type".to_Indicate.AnaVal1, BasePV := 1.0);   // "AccuS"
END_REGION
END_FUNCTION

ORGANIZATION_BLOCK "Startup"   // OB100, FBD, Startup
TITLE = "Complete Restart"
{ S7_Optimized_Access := 'TRUE' }
// stored: SetENOAutomatically false
   VAR_INPUT
      LostRetentive : Bool;   // True if retentive data are lost
      LostRTC : Bool;   // True if date and time are lost
   END_VAR
BEGIN

REGION Network 1
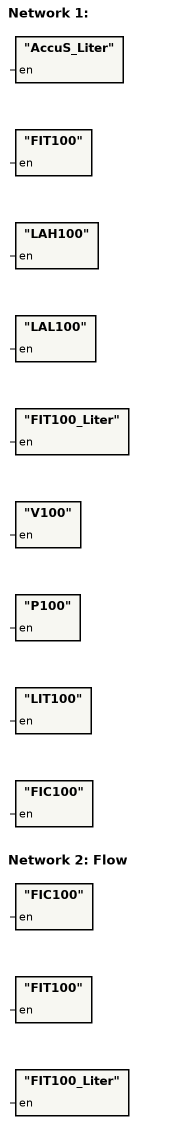
   "AccuS_Liter"();
   "FIT100"();
   "LAH100"();
   "LAL100"();
   "FIT100_Liter"();
   "V100"();
   "P100"();
   "LIT100"();
   "FIC100"();
END_REGION

REGION Network 2: Flow
   "FIC100"();
   "FIT100"();
   "FIT100_Liter"();
END_REGION

REGION Network 3: Level
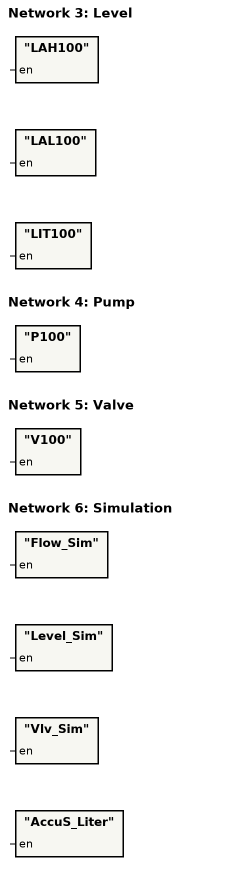
   "LAH100"();
   "LAL100"();
   "LIT100"();
END_REGION

REGION Network 4: Pump
   "P100"();
END_REGION

REGION Network 5: Valve
   "V100"();
END_REGION

REGION Network 6: Simulation
   "Flow_Sim"();
   "Level_Sim"();
   "Vlv_Sim"();
   "AccuS_Liter"();
END_REGION
END_ORGANIZATION_BLOCK

FUNCTION "ConvertToStruCm" : Void   // FC20, SCL
{ S7_Optimized_Access := 'TRUE' }
// stored: SetENOAutomatically false
   VAR_INPUT
      AnaVal1 : "AnaVal";   // Rbk
      AnaVal2 : "AnaVal";
      AnaVal3 : "AnaVal";
      DigVal1 : "DigVal";
      DigVal2 : "DigVal";
      DigVal3 : "DigVal";
      Scale : "ScaVal";   // MV_Scale
      ScaleRAW : "ScaVal_Raw";   // MV_ScaleRAW
      Unit : Int;   // MV_Unit
   END_VAR
   VAR_OUTPUT
      StruCm_Out : "StruCm";
   END_VAR
BEGIN
   #StruCm_Out.AnaVal1 := #AnaVal1;
   #StruCm_Out.AnaVal2 := #AnaVal2;
   #StruCm_Out.AnaVal3 := #AnaVal3;
   #StruCm_Out.DigVal1 := #DigVal1;
   #StruCm_Out.DigVal2 := #DigVal2;
   #StruCm_Out.DigVal3 := #DigVal3;
   #StruCm_Out.Scale := #Scale;
   #StruCm_Out.ScaleRAW := #ScaleRAW;
   #StruCm_Out.Unit := #Unit;
END_FUNCTION

FUNCTION "BoolToDigVal_1" : Void   // FC19, SCL
{ S7_Optimized_Access := 'TRUE' }
// stored: SetENOAutomatically false
   VAR_INPUT
      In : Bool;
      ST : Byte;
   END_VAR
   VAR_OUTPUT
      Out : "DigVal";
   END_VAR
BEGIN
   #Out.ST := #ST;
   #Out.Value := #In;
END_FUNCTION

DATA_BLOCK "ModuleTypePackageRevision"   // DB59
TITLE = ModuleTypePackageRevision
{ S7_Optimized_Access := 'TRUE' }
AUTHOR : Siemens AG
FAMILY : MTP
VERSION : 1.0
// The version information of the entire MTP
// stored: InstanceOfName typeMTPModuleTypePackageRevision, InstanceOfType UDT
"typeMTPModuleTypePackageRevision"
   // VAR
   //    ModuleTypePackageRevision { ExternalAccessible := 'False'; ExternalVisible := 'False'; ExternalWritable := 'False'} : String := '3.0.0';
   // END_VAR
BEGIN
END_DATA_BLOCK

DATA_BLOCK "PeaInformationLabel"   // DB14
TITLE = PeaInformationLabel
{ S7_Optimized_Access := 'TRUE' }
AUTHOR : Siemens AG
FAMILY : MTP
VERSION : 1.0
// List of product- and instance-specific information for the PEA handling within a modular plant environment.
// stored: DBAccessibleFromWebserver false, InstanceOfName typeMTPPeaInformationLabel, InstanceOfType UDT
"typeMTPPeaInformationLabel"
   // VAR
   //    AssetId : String := 'C1B54EEF-2D71-47BB-85AA-6F49015D382A';
   //    ComponentName : String := 'CleaningStationPEA';
   //    DeviceClass : String := 'CleaningStationService';
   //    DeviceHealth { ExternalWritable := 'False'} : Byte := 16#FF;
   //    DeviceManual { ExternalWritable := 'False'} : String := 'CleaningStation';
   //    DeviceRevision { ExternalWritable := 'False'} : String := '1.0.1';
   //    HardwareRevision { ExternalWritable := 'False'} : String := '1.0.1';
   //    Manufacturer { ExternalWritable := 'False'} : String := 'Siemens Presales Support';
   //    ManufacturerUri { ExternalWritable := 'False'} : String := 'https://support.industry.siemens.com/cs/de/de/view/109810699';
   //    Model { ExternalWritable := 'False'} : String := 'PresalesSupportExclusiveService';
   //    ProductCode { ExternalWritable := 'False'} : String := 'PresalesSupportPEA01';
   //    ProductInstanceUri { ExternalWritable := 'False'} : String := 'http://prtal.siemens.com/C1B54EEF-2D71-47BB-85AA-6F49015D382A';
   //    RevisionCounter { ExternalWritable := 'False'} : Int := 10;
   //    SerialNumber { ExternalWritable := 'False'} : String := 'C1B54EEF-2D71-47BB-85AA-6F49015D382A';
   //    SoftwareRevision { ExternalWritable := 'False'} : String := '2.8.0';
   // END_VAR
BEGIN
END_DATA_BLOCK

DATA_BLOCK "CMInterface_DB"   // DB27
// stored: InstanceOfName CM_Interface, InstanceOfType FB
"CM_Interface"
BEGIN
END_DATA_BLOCK

DATA_BLOCK "ConfigurationParameters_DB"   // DB32
AUTHOR : Siemens AG
FAMILY : ServiceControl
VERSION : 1.0
// stored: InstanceOfName ConfigurationParameters, InstanceOfType FB
"ConfigurationParameters"
BEGIN
   MTPBinary[0].VExt := True;
   MTPBinary[0].VOp := True;
   MTPBinary[0].VInt := True;
   MTPBinary[0].VReq := True;
   MTPBinary[0].VOut := True;
   MTPBinary[0].VState0 := 'Other PEA not co';
   MTPBinary[0].VState1 := 'Other PEA connec';
END_DATA_BLOCK

DATA_BLOCK "Dose_HMI"   // DB60
AUTHOR : Siemens AG
FAMILY : ServiceControl
VERSION : 4.0
// stored: InstanceOfName ServiceMediumParameterHMI, InstanceOfType FB
"ServiceMediumParameterHMI"
BEGIN
END_DATA_BLOCK

DATA_BLOCK "Dose_Setup"   // DB1704
TITLE = ServiceControlBlockMediumSetup
{ S7_Optimized_Access := 'TRUE'; DB_Accessible_From_OPC_UA := 'FALSE' }
AUTHOR : Siemens AG
FAMILY : ServiceControl
VERSION : 1.0
// stored: DBAccessibleFromOPCUA false, DBAccessibleFromWebserver false, InstanceOfName UDT_Service_ControlBlockMedium, InstanceOfType UDT
"UDT_Service_ControlBlockMedium"
   // VAR
   //    mode : Int := 1;
   //    stepOrder : "UDT_Service_StepOrderRawDataMedium";
   //    "step" : "UDT_Service_StepRawDataMedium";
   //    procedure : "UDT_Service_ProcedureRawDataMedium";
   //    configurationParameterData : "UDT_Service_ParameterDataMedium";
   //    processValueInData : "UDT_Service_ValueDataMedium";
   //    processValueOutData : "UDT_Service_ValueDataMedium";
   //    reportValueData : "UDT_Service_ValueDataMedium";
   //    serviceInteraction : Array[1..30] of DWord;
   //    plcGuid : String;
   //    serviceGuid : String;
   //    serviceDbNumber : Int;
   // END_VAR
BEGIN
   stepOrder.stepOrder[0].stepNumber := 0;
   stepOrder.stepOrder[1].stepNumber := 1;
   stepOrder.stepOrder[2].stepNumber := 4;
   stepOrder.stepOrder[3].stepNumber := 3;
   stepOrder.stepOrder[4].stepNumber := 5;
   stepOrder.stepOrder[5].stepNumber := 6;
   stepOrder.stepOrder[6..8].stepNumber := 2;
   stepOrder.stepOrder[9].stepNumber := 7;
   stepOrder.stepOrder[10].stepNumber := 0;
   stepOrder.stepOrder[11].stepNumber := 1;
   stepOrder.stepOrder[12].stepNumber := 4;
   stepOrder.stepOrder[13].stepNumber := 3;
   stepOrder.stepOrder[14].stepNumber := 5;
   stepOrder.stepOrder[15].stepNumber := 6;
   stepOrder.stepOrder[16..18].stepNumber := 2;
   stepOrder.stepOrder[19].stepNumber := 7;
   stepOrder.stepOrder[20].stepNumber := 0;
   stepOrder.stepOrder[21].stepNumber := 1;
   stepOrder.stepOrder[22].stepNumber := 4;
   stepOrder.stepOrder[23].stepNumber := 3;
   stepOrder.stepOrder[24].stepNumber := 5;
   stepOrder.stepOrder[25].stepNumber := 6;
   stepOrder.stepOrder[26..28].stepNumber := 2;
   stepOrder.stepOrder[29].stepNumber := 7;
   stepOrder.stepOrder[30..199].stepNumber := -1;
   stepOrder.stepOrder[0..29].stepMonitoringTime := 0;
   stepOrder.stepOrder[0..9].parameter.startIndex := 0;
   stepOrder.stepOrder[10..19].parameter.startIndex := 1;
   stepOrder.stepOrder[20..29].parameter.startIndex := -1;
   stepOrder.stepOrder[0..9].parameter.endIndex := 0;
   stepOrder.stepOrder[10..19].parameter.endIndex := 2;
   stepOrder.stepOrder[20..29].parameter.endIndex := -1;
   stepOrder.parameterIndex[0] := 16#1;
   stepOrder.parameterIndex[1] := 16#0;
   stepOrder.parameterIndex[2] := 16#1;
   "step"."step"[0].command[0] := 16#F;
   "step"."step"[1].command[0] := 16#F;
   "step"."step"[2].command[0] := 16#F;
   "step"."step"[3].command[0] := 16#3;
   "step"."step"[4].command[0] := 16#3;
   "step"."step"[5].command[0] := 16#3;
   "step"."step"[6].command[0] := 16#3;
   "step"."step"[7].command[0] := 16#0;
   "step"."step"[8].command[0] := 16#FFFF_FFFF;
   "step"."step"[9].command[0] := 16#FFFF_FFFF;
   "step"."step"[10].command[0] := 16#FFFF_FFFF;
   "step"."step"[11].command[0] := 16#FFFF_FFFF;
   "step"."step"[12].command[0] := 16#FFFF_FFFF;
   "step"."step"[13].command[0] := 16#FFFF_FFFF;
   "step"."step"[14].command[0] := 16#FFFF_FFFF;
   "step"."step"[15].command[0] := 16#FFFF_FFFF;
   "step"."step"[16].command[0] := 16#FFFF_FFFF;
   "step"."step"[17].command[0] := 16#FFFF_FFFF;
   "step"."step"[18].command[0] := 16#FFFF_FFFF;
   "step"."step"[19].command[0] := 16#FFFF_FFFF;
   "step"."step"[20].command[0] := 16#FFFF_FFFF;
   "step"."step"[21].command[0] := 16#FFFF_FFFF;
   "step"."step"[22].command[0] := 16#FFFF_FFFF;
   "step"."step"[23].command[0] := 16#FFFF_FFFF;
   "step"."step"[24].command[0] := 16#FFFF_FFFF;
   "step"."step"[25].command[0] := 16#FFFF_FFFF;
   "step"."step"[26].command[0] := 16#FFFF_FFFF;
   "step"."step"[27].command[0] := 16#FFFF_FFFF;
   "step"."step"[28].command[0] := 16#FFFF_FFFF;
   "step"."step"[29].command[0] := 16#FFFF_FFFF;
   "step"."step"[30].command[0] := 16#FFFF_FFFF;
   "step"."step"[31].command[0] := 16#FFFF_FFFF;
   "step"."step"[32].command[0] := 16#FFFF_FFFF;
   "step"."step"[33].command[0] := 16#FFFF_FFFF;
   "step"."step"[34].command[0] := 16#FFFF_FFFF;
   "step"."step"[35].command[0] := 16#FFFF_FFFF;
   "step"."step"[36].command[0] := 16#FFFF_FFFF;
   "step"."step"[37].command[0] := 16#FFFF_FFFF;
   "step"."step"[38].command[0] := 16#FFFF_FFFF;
   "step"."step"[39].command[0] := 16#FFFF_FFFF;
   "step"."step"[40].command[0] := 16#FFFF_FFFF;
   "step"."step"[41].command[0] := 16#FFFF_FFFF;
   "step"."step"[42].command[0] := 16#FFFF_FFFF;
   "step"."step"[43].command[0] := 16#FFFF_FFFF;
   "step"."step"[44].command[0] := 16#FFFF_FFFF;
   "step"."step"[45].command[0] := 16#FFFF_FFFF;
   "step"."step"[46].command[0] := 16#FFFF_FFFF;
   "step"."step"[47].command[0] := 16#FFFF_FFFF;
   "step"."step"[48].command[0] := 16#FFFF_FFFF;
   "step"."step"[49].command[0] := 16#FFFF_FFFF;
   "step"."step"[50].command[0] := 16#FFFF_FFFF;
   "step"."step"[51].command[0] := 16#FFFF_FFFF;
   "step"."step"[52].command[0] := 16#FFFF_FFFF;
   "step"."step"[53].command[0] := 16#FFFF_FFFF;
   "step"."step"[54].command[0] := 16#FFFF_FFFF;
   "step"."step"[55].command[0] := 16#FFFF_FFFF;
   "step"."step"[56].command[0] := 16#FFFF_FFFF;
   "step"."step"[57].command[0] := 16#FFFF_FFFF;
   "step"."step"[58].command[0] := 16#FFFF_FFFF;
   "step"."step"[59].command[0] := 16#FFFF_FFFF;
   "step"."step"[60].command[0] := 16#FFFF_FFFF;
   "step"."step"[61].command[0] := 16#FFFF_FFFF;
   "step"."step"[62].command[0] := 16#FFFF_FFFF;
   "step"."step"[63].command[0] := 16#FFFF_FFFF;
   "step"."step"[64].command[0] := 16#FFFF_FFFF;
   "step"."step"[65].command[0] := 16#FFFF_FFFF;
   "step"."step"[66].command[0] := 16#FFFF_FFFF;
   "step"."step"[67].command[0] := 16#FFFF_FFFF;
   "step"."step"[68].command[0] := 16#FFFF_FFFF;
   "step"."step"[69].command[0] := 16#FFFF_FFFF;
   "step"."step"[70].command[0] := 16#FFFF_FFFF;
   "step"."step"[71].command[0] := 16#FFFF_FFFF;
   "step"."step"[72].command[0] := 16#FFFF_FFFF;
   "step"."step"[73].command[0] := 16#FFFF_FFFF;
   "step"."step"[74].command[0] := 16#FFFF_FFFF;
   "step"."step"[75].command[0] := 16#FFFF_FFFF;
   "step"."step"[76].command[0] := 16#FFFF_FFFF;
   "step"."step"[77].command[0] := 16#FFFF_FFFF;
   "step"."step"[78].command[0] := 16#FFFF_FFFF;
   "step"."step"[79].command[0] := 16#FFFF_FFFF;
   "step"."step"[80].command[0] := 16#FFFF_FFFF;
   "step"."step"[81].command[0] := 16#FFFF_FFFF;
   "step"."step"[82].command[0] := 16#FFFF_FFFF;
   "step"."step"[83].command[0] := 16#FFFF_FFFF;
   "step"."step"[84].command[0] := 16#FFFF_FFFF;
   "step"."step"[85].command[0] := 16#FFFF_FFFF;
   "step"."step"[86].command[0] := 16#FFFF_FFFF;
   "step"."step"[87].command[0] := 16#FFFF_FFFF;
   "step"."step"[88].command[0] := 16#FFFF_FFFF;
   "step"."step"[89].command[0] := 16#FFFF_FFFF;
   "step"."step"[90].command[0] := 16#FFFF_FFFF;
   "step"."step"[91].command[0] := 16#FFFF_FFFF;
   "step"."step"[92].command[0] := 16#FFFF_FFFF;
   "step"."step"[93].command[0] := 16#FFFF_FFFF;
   "step"."step"[94].command[0] := 16#FFFF_FFFF;
   "step"."step"[95].command[0] := 16#FFFF_FFFF;
   "step"."step"[96].command[0] := 16#FFFF_FFFF;
   "step"."step"[97].command[0] := 16#FFFF_FFFF;
   "step"."step"[98].command[0] := 16#FFFF_FFFF;
   "step"."step"[99].command[0] := 16#FFFF_FFFF;
   "step"."step"[0].force[0] := 16#F;
   "step"."step"[1].force[0] := 16#F;
   "step"."step"[2].force[0] := 16#F;
   "step"."step"[3].force[0] := 16#3;
   "step"."step"[4].force[0] := 16#3;
   "step"."step"[5].force[0] := 16#3;
   "step"."step"[6].force[0] := 16#3;
   "step"."step"[7].force[0] := 16#0;
   "step"."step"[8].force[0] := 16#FFFF_FFFF;
   "step"."step"[9].force[0] := 16#FFFF_FFFF;
   "step"."step"[10].force[0] := 16#FFFF_FFFF;
   "step"."step"[11].force[0] := 16#FFFF_FFFF;
   "step"."step"[12].force[0] := 16#FFFF_FFFF;
   "step"."step"[13].force[0] := 16#FFFF_FFFF;
   "step"."step"[14].force[0] := 16#FFFF_FFFF;
   "step"."step"[15].force[0] := 16#FFFF_FFFF;
   "step"."step"[16].force[0] := 16#FFFF_FFFF;
   "step"."step"[17].force[0] := 16#FFFF_FFFF;
   "step"."step"[18].force[0] := 16#FFFF_FFFF;
   "step"."step"[19].force[0] := 16#FFFF_FFFF;
   "step"."step"[20].force[0] := 16#FFFF_FFFF;
   "step"."step"[21].force[0] := 16#FFFF_FFFF;
   "step"."step"[22].force[0] := 16#FFFF_FFFF;
   "step"."step"[23].force[0] := 16#FFFF_FFFF;
   "step"."step"[24].force[0] := 16#FFFF_FFFF;
   "step"."step"[25].force[0] := 16#FFFF_FFFF;
   "step"."step"[26].force[0] := 16#FFFF_FFFF;
   "step"."step"[27].force[0] := 16#FFFF_FFFF;
   "step"."step"[28].force[0] := 16#FFFF_FFFF;
   "step"."step"[29].force[0] := 16#FFFF_FFFF;
   "step"."step"[30].force[0] := 16#FFFF_FFFF;
   "step"."step"[31].force[0] := 16#FFFF_FFFF;
   "step"."step"[32].force[0] := 16#FFFF_FFFF;
   "step"."step"[33].force[0] := 16#FFFF_FFFF;
   "step"."step"[34].force[0] := 16#FFFF_FFFF;
   "step"."step"[35].force[0] := 16#FFFF_FFFF;
   "step"."step"[36].force[0] := 16#FFFF_FFFF;
   "step"."step"[37].force[0] := 16#FFFF_FFFF;
   "step"."step"[38].force[0] := 16#FFFF_FFFF;
   "step"."step"[39].force[0] := 16#FFFF_FFFF;
   "step"."step"[40].force[0] := 16#FFFF_FFFF;
   "step"."step"[41].force[0] := 16#FFFF_FFFF;
   "step"."step"[42].force[0] := 16#FFFF_FFFF;
   "step"."step"[43].force[0] := 16#FFFF_FFFF;
   "step"."step"[44].force[0] := 16#FFFF_FFFF;
   "step"."step"[45].force[0] := 16#FFFF_FFFF;
   "step"."step"[46].force[0] := 16#FFFF_FFFF;
   "step"."step"[47].force[0] := 16#FFFF_FFFF;
   "step"."step"[48].force[0] := 16#FFFF_FFFF;
   "step"."step"[49].force[0] := 16#FFFF_FFFF;
   "step"."step"[50].force[0] := 16#FFFF_FFFF;
   "step"."step"[51].force[0] := 16#FFFF_FFFF;
   "step"."step"[52].force[0] := 16#FFFF_FFFF;
   "step"."step"[53].force[0] := 16#FFFF_FFFF;
   "step"."step"[54].force[0] := 16#FFFF_FFFF;
   "step"."step"[55].force[0] := 16#FFFF_FFFF;
   "step"."step"[56].force[0] := 16#FFFF_FFFF;
   "step"."step"[57].force[0] := 16#FFFF_FFFF;
   "step"."step"[58].force[0] := 16#FFFF_FFFF;
   "step"."step"[59].force[0] := 16#FFFF_FFFF;
   "step"."step"[60].force[0] := 16#FFFF_FFFF;
   "step"."step"[61].force[0] := 16#FFFF_FFFF;
   "step"."step"[62].force[0] := 16#FFFF_FFFF;
   "step"."step"[63].force[0] := 16#FFFF_FFFF;
   "step"."step"[64].force[0] := 16#FFFF_FFFF;
   "step"."step"[65].force[0] := 16#FFFF_FFFF;
   "step"."step"[66].force[0] := 16#FFFF_FFFF;
   "step"."step"[67].force[0] := 16#FFFF_FFFF;
   "step"."step"[68].force[0] := 16#FFFF_FFFF;
   "step"."step"[69].force[0] := 16#FFFF_FFFF;
   "step"."step"[70].force[0] := 16#FFFF_FFFF;
   "step"."step"[71].force[0] := 16#FFFF_FFFF;
   "step"."step"[72].force[0] := 16#FFFF_FFFF;
   "step"."step"[73].force[0] := 16#FFFF_FFFF;
   "step"."step"[74].force[0] := 16#FFFF_FFFF;
   "step"."step"[75].force[0] := 16#FFFF_FFFF;
   "step"."step"[76].force[0] := 16#FFFF_FFFF;
   "step"."step"[77].force[0] := 16#FFFF_FFFF;
   "step"."step"[78].force[0] := 16#FFFF_FFFF;
   "step"."step"[79].force[0] := 16#FFFF_FFFF;
   "step"."step"[80].force[0] := 16#FFFF_FFFF;
   "step"."step"[81].force[0] := 16#FFFF_FFFF;
   "step"."step"[82].force[0] := 16#FFFF_FFFF;
   "step"."step"[83].force[0] := 16#FFFF_FFFF;
   "step"."step"[84].force[0] := 16#FFFF_FFFF;
   "step"."step"[85].force[0] := 16#FFFF_FFFF;
   "step"."step"[86].force[0] := 16#FFFF_FFFF;
   "step"."step"[87].force[0] := 16#FFFF_FFFF;
   "step"."step"[88].force[0] := 16#FFFF_FFFF;
   "step"."step"[89].force[0] := 16#FFFF_FFFF;
   "step"."step"[90].force[0] := 16#FFFF_FFFF;
   "step"."step"[91].force[0] := 16#FFFF_FFFF;
   "step"."step"[92].force[0] := 16#FFFF_FFFF;
   "step"."step"[93].force[0] := 16#FFFF_FFFF;
   "step"."step"[94].force[0] := 16#FFFF_FFFF;
   "step"."step"[95].force[0] := 16#FFFF_FFFF;
   "step"."step"[96].force[0] := 16#FFFF_FFFF;
   "step"."step"[97].force[0] := 16#FFFF_FFFF;
   "step"."step"[98].force[0] := 16#FFFF_FFFF;
   "step"."step"[99].force[0] := 16#FFFF_FFFF;
   "step"."step"[0].check[0] := 16#F;
   "step"."step"[1].check[0] := 16#F;
   "step"."step"[2].check[0] := 16#F;
   "step"."step"[3].check[0] := 16#3;
   "step"."step"[4].check[0] := 16#3;
   "step"."step"[5].check[0] := 16#3;
   "step"."step"[6].check[0] := 16#0;
   "step"."step"[7].check[0] := 16#0;
   "step"."step"[8].check[0] := 16#FFFF_FFFF;
   "step"."step"[9].check[0] := 16#FFFF_FFFF;
   "step"."step"[10].check[0] := 16#FFFF_FFFF;
   "step"."step"[11].check[0] := 16#FFFF_FFFF;
   "step"."step"[12].check[0] := 16#FFFF_FFFF;
   "step"."step"[13].check[0] := 16#FFFF_FFFF;
   "step"."step"[14].check[0] := 16#FFFF_FFFF;
   "step"."step"[15].check[0] := 16#FFFF_FFFF;
   "step"."step"[16].check[0] := 16#FFFF_FFFF;
   "step"."step"[17].check[0] := 16#FFFF_FFFF;
   "step"."step"[18].check[0] := 16#FFFF_FFFF;
   "step"."step"[19].check[0] := 16#FFFF_FFFF;
   "step"."step"[20].check[0] := 16#FFFF_FFFF;
   "step"."step"[21].check[0] := 16#FFFF_FFFF;
   "step"."step"[22].check[0] := 16#FFFF_FFFF;
   "step"."step"[23].check[0] := 16#FFFF_FFFF;
   "step"."step"[24].check[0] := 16#FFFF_FFFF;
   "step"."step"[25].check[0] := 16#FFFF_FFFF;
   "step"."step"[26].check[0] := 16#FFFF_FFFF;
   "step"."step"[27].check[0] := 16#FFFF_FFFF;
   "step"."step"[28].check[0] := 16#FFFF_FFFF;
   "step"."step"[29].check[0] := 16#FFFF_FFFF;
   "step"."step"[30].check[0] := 16#FFFF_FFFF;
   "step"."step"[31].check[0] := 16#FFFF_FFFF;
   "step"."step"[32].check[0] := 16#FFFF_FFFF;
   "step"."step"[33].check[0] := 16#FFFF_FFFF;
   "step"."step"[34].check[0] := 16#FFFF_FFFF;
   "step"."step"[35].check[0] := 16#FFFF_FFFF;
   "step"."step"[36].check[0] := 16#FFFF_FFFF;
   "step"."step"[37].check[0] := 16#FFFF_FFFF;
   "step"."step"[38].check[0] := 16#FFFF_FFFF;
   "step"."step"[39].check[0] := 16#FFFF_FFFF;
   "step"."step"[40].check[0] := 16#FFFF_FFFF;
   "step"."step"[41].check[0] := 16#FFFF_FFFF;
   "step"."step"[42].check[0] := 16#FFFF_FFFF;
   "step"."step"[43].check[0] := 16#FFFF_FFFF;
   "step"."step"[44].check[0] := 16#FFFF_FFFF;
   "step"."step"[45].check[0] := 16#FFFF_FFFF;
   "step"."step"[46].check[0] := 16#FFFF_FFFF;
   "step"."step"[47].check[0] := 16#FFFF_FFFF;
   "step"."step"[48].check[0] := 16#FFFF_FFFF;
   "step"."step"[49].check[0] := 16#FFFF_FFFF;
   "step"."step"[50].check[0] := 16#FFFF_FFFF;
   "step"."step"[51].check[0] := 16#FFFF_FFFF;
   "step"."step"[52].check[0] := 16#FFFF_FFFF;
   "step"."step"[53].check[0] := 16#FFFF_FFFF;
   "step"."step"[54].check[0] := 16#FFFF_FFFF;
   "step"."step"[55].check[0] := 16#FFFF_FFFF;
   "step"."step"[56].check[0] := 16#FFFF_FFFF;
   "step"."step"[57].check[0] := 16#FFFF_FFFF;
   "step"."step"[58].check[0] := 16#FFFF_FFFF;
   "step"."step"[59].check[0] := 16#FFFF_FFFF;
   "step"."step"[60].check[0] := 16#FFFF_FFFF;
   "step"."step"[61].check[0] := 16#FFFF_FFFF;
   "step"."step"[62].check[0] := 16#FFFF_FFFF;
   "step"."step"[63].check[0] := 16#FFFF_FFFF;
   "step"."step"[64].check[0] := 16#FFFF_FFFF;
   "step"."step"[65].check[0] := 16#FFFF_FFFF;
   "step"."step"[66].check[0] := 16#FFFF_FFFF;
   "step"."step"[67].check[0] := 16#FFFF_FFFF;
   "step"."step"[68].check[0] := 16#FFFF_FFFF;
   "step"."step"[69].check[0] := 16#FFFF_FFFF;
   "step"."step"[70].check[0] := 16#FFFF_FFFF;
   "step"."step"[71].check[0] := 16#FFFF_FFFF;
   "step"."step"[72].check[0] := 16#FFFF_FFFF;
   "step"."step"[73].check[0] := 16#FFFF_FFFF;
   "step"."step"[74].check[0] := 16#FFFF_FFFF;
   "step"."step"[75].check[0] := 16#FFFF_FFFF;
   "step"."step"[76].check[0] := 16#FFFF_FFFF;
   "step"."step"[77].check[0] := 16#FFFF_FFFF;
   "step"."step"[78].check[0] := 16#FFFF_FFFF;
   "step"."step"[79].check[0] := 16#FFFF_FFFF;
   "step"."step"[80].check[0] := 16#FFFF_FFFF;
   "step"."step"[81].check[0] := 16#FFFF_FFFF;
   "step"."step"[82].check[0] := 16#FFFF_FFFF;
   "step"."step"[83].check[0] := 16#FFFF_FFFF;
   "step"."step"[84].check[0] := 16#FFFF_FFFF;
   "step"."step"[85].check[0] := 16#FFFF_FFFF;
   "step"."step"[86].check[0] := 16#FFFF_FFFF;
   "step"."step"[87].check[0] := 16#FFFF_FFFF;
   "step"."step"[88].check[0] := 16#FFFF_FFFF;
   "step"."step"[89].check[0] := 16#FFFF_FFFF;
   "step"."step"[90].check[0] := 16#FFFF_FFFF;
   "step"."step"[91].check[0] := 16#FFFF_FFFF;
   "step"."step"[92].check[0] := 16#FFFF_FFFF;
   "step"."step"[93].check[0] := 16#FFFF_FFFF;
   "step"."step"[94].check[0] := 16#FFFF_FFFF;
   "step"."step"[95].check[0] := 16#FFFF_FFFF;
   "step"."step"[96].check[0] := 16#FFFF_FFFF;
   "step"."step"[97].check[0] := 16#FFFF_FFFF;
   "step"."step"[98].check[0] := 16#FFFF_FFFF;
   "step"."step"[99].check[0] := 16#FFFF_FFFF;
   "step"."step"[0]."or"[0] := 16#0;
   "step"."step"[1]."or"[0] := 16#0;
   "step"."step"[2]."or"[0] := 16#0;
   "step"."step"[3]."or"[0] := 16#0;
   "step"."step"[4]."or"[0] := 16#0;
   "step"."step"[5]."or"[0] := 16#0;
   "step"."step"[6]."or"[0] := 16#0;
   "step"."step"[7]."or"[0] := 16#0;
   "step"."step"[8]."or"[0] := 16#FFFF_FFFF;
   "step"."step"[9]."or"[0] := 16#FFFF_FFFF;
   "step"."step"[10]."or"[0] := 16#FFFF_FFFF;
   "step"."step"[11]."or"[0] := 16#FFFF_FFFF;
   "step"."step"[12]."or"[0] := 16#FFFF_FFFF;
   "step"."step"[13]."or"[0] := 16#FFFF_FFFF;
   "step"."step"[14]."or"[0] := 16#FFFF_FFFF;
   "step"."step"[15]."or"[0] := 16#FFFF_FFFF;
   "step"."step"[16]."or"[0] := 16#FFFF_FFFF;
   "step"."step"[17]."or"[0] := 16#FFFF_FFFF;
   "step"."step"[18]."or"[0] := 16#FFFF_FFFF;
   "step"."step"[19]."or"[0] := 16#FFFF_FFFF;
   "step"."step"[20]."or"[0] := 16#FFFF_FFFF;
   "step"."step"[21]."or"[0] := 16#FFFF_FFFF;
   "step"."step"[22]."or"[0] := 16#FFFF_FFFF;
   "step"."step"[23]."or"[0] := 16#FFFF_FFFF;
   "step"."step"[24]."or"[0] := 16#FFFF_FFFF;
   "step"."step"[25]."or"[0] := 16#FFFF_FFFF;
   "step"."step"[26]."or"[0] := 16#FFFF_FFFF;
   "step"."step"[27]."or"[0] := 16#FFFF_FFFF;
   "step"."step"[28]."or"[0] := 16#FFFF_FFFF;
   "step"."step"[29]."or"[0] := 16#FFFF_FFFF;
   "step"."step"[30]."or"[0] := 16#FFFF_FFFF;
   "step"."step"[31]."or"[0] := 16#FFFF_FFFF;
   "step"."step"[32]."or"[0] := 16#FFFF_FFFF;
   "step"."step"[33]."or"[0] := 16#FFFF_FFFF;
   "step"."step"[34]."or"[0] := 16#FFFF_FFFF;
   "step"."step"[35]."or"[0] := 16#FFFF_FFFF;
   "step"."step"[36]."or"[0] := 16#FFFF_FFFF;
   "step"."step"[37]."or"[0] := 16#FFFF_FFFF;
   "step"."step"[38]."or"[0] := 16#FFFF_FFFF;
   "step"."step"[39]."or"[0] := 16#FFFF_FFFF;
   "step"."step"[40]."or"[0] := 16#FFFF_FFFF;
   "step"."step"[41]."or"[0] := 16#FFFF_FFFF;
   "step"."step"[42]."or"[0] := 16#FFFF_FFFF;
   "step"."step"[43]."or"[0] := 16#FFFF_FFFF;
   "step"."step"[44]."or"[0] := 16#FFFF_FFFF;
   "step"."step"[45]."or"[0] := 16#FFFF_FFFF;
   "step"."step"[46]."or"[0] := 16#FFFF_FFFF;
   "step"."step"[47]."or"[0] := 16#FFFF_FFFF;
   "step"."step"[48]."or"[0] := 16#FFFF_FFFF;
   "step"."step"[49]."or"[0] := 16#FFFF_FFFF;
   "step"."step"[50]."or"[0] := 16#FFFF_FFFF;
   "step"."step"[51]."or"[0] := 16#FFFF_FFFF;
   "step"."step"[52]."or"[0] := 16#FFFF_FFFF;
   "step"."step"[53]."or"[0] := 16#FFFF_FFFF;
   "step"."step"[54]."or"[0] := 16#FFFF_FFFF;
   "step"."step"[55]."or"[0] := 16#FFFF_FFFF;
   "step"."step"[56]."or"[0] := 16#FFFF_FFFF;
   "step"."step"[57]."or"[0] := 16#FFFF_FFFF;
   "step"."step"[58]."or"[0] := 16#FFFF_FFFF;
   "step"."step"[59]."or"[0] := 16#FFFF_FFFF;
   "step"."step"[60]."or"[0] := 16#FFFF_FFFF;
   "step"."step"[61]."or"[0] := 16#FFFF_FFFF;
   "step"."step"[62]."or"[0] := 16#FFFF_FFFF;
   "step"."step"[63]."or"[0] := 16#FFFF_FFFF;
   "step"."step"[64]."or"[0] := 16#FFFF_FFFF;
   "step"."step"[65]."or"[0] := 16#FFFF_FFFF;
   "step"."step"[66]."or"[0] := 16#FFFF_FFFF;
   "step"."step"[67]."or"[0] := 16#FFFF_FFFF;
   "step"."step"[68]."or"[0] := 16#FFFF_FFFF;
   "step"."step"[69]."or"[0] := 16#FFFF_FFFF;
   "step"."step"[70]."or"[0] := 16#FFFF_FFFF;
   "step"."step"[71]."or"[0] := 16#FFFF_FFFF;
   "step"."step"[72]."or"[0] := 16#FFFF_FFFF;
   "step"."step"[73]."or"[0] := 16#FFFF_FFFF;
   "step"."step"[74]."or"[0] := 16#FFFF_FFFF;
   "step"."step"[75]."or"[0] := 16#FFFF_FFFF;
   "step"."step"[76]."or"[0] := 16#FFFF_FFFF;
   "step"."step"[77]."or"[0] := 16#FFFF_FFFF;
   "step"."step"[78]."or"[0] := 16#FFFF_FFFF;
   "step"."step"[79]."or"[0] := 16#FFFF_FFFF;
   "step"."step"[80]."or"[0] := 16#FFFF_FFFF;
   "step"."step"[81]."or"[0] := 16#FFFF_FFFF;
   "step"."step"[82]."or"[0] := 16#FFFF_FFFF;
   "step"."step"[83]."or"[0] := 16#FFFF_FFFF;
   "step"."step"[84]."or"[0] := 16#FFFF_FFFF;
   "step"."step"[85]."or"[0] := 16#FFFF_FFFF;
   "step"."step"[86]."or"[0] := 16#FFFF_FFFF;
   "step"."step"[87]."or"[0] := 16#FFFF_FFFF;
   "step"."step"[88]."or"[0] := 16#FFFF_FFFF;
   "step"."step"[89]."or"[0] := 16#FFFF_FFFF;
   "step"."step"[90]."or"[0] := 16#FFFF_FFFF;
   "step"."step"[91]."or"[0] := 16#FFFF_FFFF;
   "step"."step"[92]."or"[0] := 16#FFFF_FFFF;
   "step"."step"[93]."or"[0] := 16#FFFF_FFFF;
   "step"."step"[94]."or"[0] := 16#FFFF_FFFF;
   "step"."step"[95]."or"[0] := 16#FFFF_FFFF;
   "step"."step"[96]."or"[0] := 16#FFFF_FFFF;
   "step"."step"[97]."or"[0] := 16#FFFF_FFFF;
   "step"."step"[98]."or"[0] := 16#FFFF_FFFF;
   "step"."step"[99]."or"[0] := 16#FFFF_FFFF;
   "step".parameterDefinition[0].indexMTP := 0;
   "step".parameterDefinition[1].indexMTP := 1;
   "step".parameterDefinition[0].indexIO := 0;
   "step".parameterDefinition[1].indexIO := 1;
   "step".parameterDefinition[0..1]."type" := 1;
   "step".parameterDefinition[0..1].controlModule := 16#0;
   "step".parameterDefinition[2..31].controlModule := 16#FF;
   procedure.procedure[0..2].Procedure.IsSelfCompleting := True;
   procedure.procedure[3..15].Procedure.IsSelfCompleting := False;
   procedure.procedure[0].Procedure.ProcedureID := 16#1;
   procedure.procedure[1].Procedure.ProcedureID := 16#2;
   procedure.procedure[2].Procedure.ProcedureID := 16#3;
   procedure.procedure[3..15].Procedure.ProcedureID := 16#0;
   procedure.procedure[0..15].Procedure.IsDefault := False;
   procedure.procedure[0].StateTransient.starting.startIndex := 0;
   procedure.procedure[1].StateTransient.starting.startIndex := 10;
   procedure.procedure[2].StateTransient.starting.startIndex := 20;
   procedure.procedure[3..15].StateTransient.starting.startIndex := -1;
   procedure.procedure[0].StateTransient.starting.endIndex := 0;
   procedure.procedure[1].StateTransient.starting.endIndex := 10;
   procedure.procedure[2].StateTransient.starting.endIndex := 20;
   procedure.procedure[3..15].StateTransient.starting.endIndex := -1;
   procedure.procedure[0].StateTransient.running.startIndex := 1;
   procedure.procedure[1].StateTransient.running.startIndex := 11;
   procedure.procedure[2].StateTransient.running.startIndex := 21;
   procedure.procedure[3..15].StateTransient.running.startIndex := -1;
   procedure.procedure[0].StateTransient.running.endIndex := 1;
   procedure.procedure[1].StateTransient.running.endIndex := 11;
   procedure.procedure[2].StateTransient.running.endIndex := 21;
   procedure.procedure[3..15].StateTransient.running.endIndex := -1;
   procedure.procedure[0].StateTransient.holding.startIndex := 2;
   procedure.procedure[1].StateTransient.holding.startIndex := 12;
   procedure.procedure[2].StateTransient.holding.startIndex := 22;
   procedure.procedure[3..15].StateTransient.holding.startIndex := -1;
   procedure.procedure[0].StateTransient.holding.endIndex := 2;
   procedure.procedure[1].StateTransient.holding.endIndex := 12;
   procedure.procedure[2].StateTransient.holding.endIndex := 22;
   procedure.procedure[3..15].StateTransient.holding.endIndex := -1;
   procedure.procedure[0].StateTransient.unholding.startIndex := 3;
   procedure.procedure[1].StateTransient.unholding.startIndex := 13;
   procedure.procedure[2].StateTransient.unholding.startIndex := 23;
   procedure.procedure[3..15].StateTransient.unholding.startIndex := -1;
   procedure.procedure[0].StateTransient.unholding.endIndex := 3;
   procedure.procedure[1].StateTransient.unholding.endIndex := 13;
   procedure.procedure[2].StateTransient.unholding.endIndex := 23;
   procedure.procedure[3..15].StateTransient.unholding.endIndex := -1;
   procedure.procedure[0].StateTransient.pausing.startIndex := 4;
   procedure.procedure[1].StateTransient.pausing.startIndex := 14;
   procedure.procedure[2].StateTransient.pausing.startIndex := 24;
   procedure.procedure[3..15].StateTransient.pausing.startIndex := -1;
   procedure.procedure[0].StateTransient.pausing.endIndex := 4;
   procedure.procedure[1].StateTransient.pausing.endIndex := 14;
   procedure.procedure[2].StateTransient.pausing.endIndex := 24;
   procedure.procedure[3..15].StateTransient.pausing.endIndex := -1;
   procedure.procedure[0].StateTransient.resuming.startIndex := 5;
   procedure.procedure[1].StateTransient.resuming.startIndex := 15;
   procedure.procedure[2].StateTransient.resuming.startIndex := 25;
   procedure.procedure[3..15].StateTransient.resuming.startIndex := -1;
   procedure.procedure[0].StateTransient.resuming.endIndex := 5;
   procedure.procedure[1].StateTransient.resuming.endIndex := 15;
   procedure.procedure[2].StateTransient.resuming.endIndex := 25;
   procedure.procedure[3..15].StateTransient.resuming.endIndex := -1;
   procedure.procedure[0].StateTransient.completing.startIndex := 6;
   procedure.procedure[1].StateTransient.completing.startIndex := 16;
   procedure.procedure[2].StateTransient.completing.startIndex := 26;
   procedure.procedure[3..15].StateTransient.completing.startIndex := -1;
   procedure.procedure[0].StateTransient.completing.endIndex := 6;
   procedure.procedure[1].StateTransient.completing.endIndex := 16;
   procedure.procedure[2].StateTransient.completing.endIndex := 26;
   procedure.procedure[3..15].StateTransient.completing.endIndex := -1;
   procedure.procedure[0].StateTransient.stopping.startIndex := 7;
   procedure.procedure[1].StateTransient.stopping.startIndex := 17;
   procedure.procedure[2].StateTransient.stopping.startIndex := 27;
   procedure.procedure[3..15].StateTransient.stopping.startIndex := -1;
   procedure.procedure[0].StateTransient.stopping.endIndex := 7;
   procedure.procedure[1].StateTransient.stopping.endIndex := 17;
   procedure.procedure[2].StateTransient.stopping.endIndex := 27;
   procedure.procedure[3..15].StateTransient.stopping.endIndex := -1;
   procedure.procedure[0].StateTransient.aborting.startIndex := 8;
   procedure.procedure[1].StateTransient.aborting.startIndex := 18;
   procedure.procedure[2].StateTransient.aborting.startIndex := 28;
   procedure.procedure[3..15].StateTransient.aborting.startIndex := -1;
   procedure.procedure[0].StateTransient.aborting.endIndex := 8;
   procedure.procedure[1].StateTransient.aborting.endIndex := 18;
   procedure.procedure[2].StateTransient.aborting.endIndex := 28;
   procedure.procedure[3..15].StateTransient.aborting.endIndex := -1;
   procedure.procedure[0].StateTransient.resetting.startIndex := 9;
   procedure.procedure[1].StateTransient.resetting.startIndex := 19;
   procedure.procedure[2].StateTransient.resetting.startIndex := 29;
   procedure.procedure[3..15].StateTransient.resetting.startIndex := -1;
   procedure.procedure[0].StateTransient.resetting.endIndex := 9;
   procedure.procedure[1].StateTransient.resetting.endIndex := 19;
   procedure.procedure[2].StateTransient.resetting.endIndex := 29;
   procedure.procedure[3..15].StateTransient.resetting.endIndex := -1;
   procedure.procedure[0].ProcedureReportMap[0] := 16#1;
   procedure.procedure[1].ProcedureReportMap[0] := 16#1;
   procedure.procedure[2].ProcedureReportMap[0] := 16#1;
   procedure.procedure[3].ProcedureReportMap[0] := 16#0;
   procedure.procedure[4].ProcedureReportMap[0] := 16#0;
   procedure.procedure[5].ProcedureReportMap[0] := 16#0;
   procedure.procedure[6].ProcedureReportMap[0] := 16#0;
   procedure.procedure[7].ProcedureReportMap[0] := 16#0;
   procedure.procedure[8].ProcedureReportMap[0] := 16#0;
   procedure.procedure[9].ProcedureReportMap[0] := 16#0;
   procedure.procedure[10].ProcedureReportMap[0] := 16#0;
   procedure.procedure[11].ProcedureReportMap[0] := 16#0;
   procedure.procedure[12].ProcedureReportMap[0] := 16#0;
   procedure.procedure[13].ProcedureReportMap[0] := 16#0;
   procedure.procedure[14].ProcedureReportMap[0] := 16#0;
   procedure.procedure[15].ProcedureReportMap[0] := 16#0;
   procedure.procedure[0].ProcedureProcessInMap[0] := 16#3;
   procedure.procedure[1].ProcedureProcessInMap[0] := 16#3;
   procedure.procedure[2].ProcedureProcessInMap[0] := 16#3;
   procedure.procedure[3].ProcedureProcessInMap[0] := 16#0;
   procedure.procedure[4].ProcedureProcessInMap[0] := 16#0;
   procedure.procedure[5].ProcedureProcessInMap[0] := 16#0;
   procedure.procedure[6].ProcedureProcessInMap[0] := 16#0;
   procedure.procedure[7].ProcedureProcessInMap[0] := 16#0;
   procedure.procedure[8].ProcedureProcessInMap[0] := 16#0;
   procedure.procedure[9].ProcedureProcessInMap[0] := 16#0;
   procedure.procedure[10].ProcedureProcessInMap[0] := 16#0;
   procedure.procedure[11].ProcedureProcessInMap[0] := 16#0;
   procedure.procedure[12].ProcedureProcessInMap[0] := 16#0;
   procedure.procedure[13].ProcedureProcessInMap[0] := 16#0;
   procedure.procedure[14].ProcedureProcessInMap[0] := 16#0;
   procedure.procedure[15].ProcedureProcessInMap[0] := 16#0;
   procedure.procedure[0].ProcedureProcessOutMap[0] := 16#1;
   procedure.procedure[1].ProcedureProcessOutMap[0] := 16#1;
   procedure.procedure[2].ProcedureProcessOutMap[0] := 16#1;
   procedure.procedure[3].ProcedureProcessOutMap[0] := 16#0;
   procedure.procedure[4].ProcedureProcessOutMap[0] := 16#0;
   procedure.procedure[5].ProcedureProcessOutMap[0] := 16#0;
   procedure.procedure[6].ProcedureProcessOutMap[0] := 16#0;
   procedure.procedure[7].ProcedureProcessOutMap[0] := 16#0;
   procedure.procedure[8].ProcedureProcessOutMap[0] := 16#0;
   procedure.procedure[9].ProcedureProcessOutMap[0] := 16#0;
   procedure.procedure[10].ProcedureProcessOutMap[0] := 16#0;
   procedure.procedure[11].ProcedureProcessOutMap[0] := 16#0;
   procedure.procedure[12].ProcedureProcessOutMap[0] := 16#0;
   procedure.procedure[13].ProcedureProcessOutMap[0] := 16#0;
   procedure.procedure[14].ProcedureProcessOutMap[0] := 16#0;
   procedure.procedure[15].ProcedureProcessOutMap[0] := 16#0;
   configurationParameterData.used[0] := 16#1;
   configurationParameterData.definition[0].indexMTP := 0;
   configurationParameterData.definition[0].indexIO := 0;
   configurationParameterData.definition[0]."type" := 3;
   configurationParameterData.definition[0].controlModule := 16#0;
   configurationParameterData.definition[1..31].controlModule := 16#FF;
   processValueInData.used[0] := 16#1;
   processValueInData.definition[0..1].indexMTP := 0;
   processValueInData.definition[0..1].indexIO := 0;
   processValueInData.definition[0]."type" := 1;
   processValueInData.definition[1]."type" := 3;
   processValueInData.definition[0..1].controlModule := 16#0;
   processValueInData.definition[2..31].controlModule := 16#FF;
   processValueOutData.used[0] := 16#1;
   processValueOutData.definition[0].indexMTP := 0;
   processValueOutData.definition[0].indexIO := 0;
   processValueOutData.definition[0]."type" := 1;
   processValueOutData.definition[0].controlModule := 16#0;
   processValueOutData.definition[1..31].controlModule := 16#FF;
   reportValueData.used[0] := 16#1;
   reportValueData.definition[0].indexMTP := 0;
   reportValueData.definition[1].indexMTP := 1;
   reportValueData.definition[0].indexIO := 0;
   reportValueData.definition[1].indexIO := 1;
   reportValueData.definition[0..1]."type" := 1;
   reportValueData.definition[0].controlModule := 16#0;
   reportValueData.definition[1..31].controlModule := 16#FF;
   serviceInteraction[1] := 16#1;
   serviceInteraction[2..30] := 16#0;
END_DATA_BLOCK

DATA_BLOCK "ProcedureParameters_DB"   // DB33
AUTHOR : Siemens AG
FAMILY : ServiceControl
VERSION : 1.0
// stored: InstanceOfName ProcedureParameters, InstanceOfType FB
"ProcedureParameters"
BEGIN
   MTPAnalog[0..2].Sync := True;
   MTPAnalog[0].VExt := 25.0;
   MTPAnalog[1].VExt := 1000.0;
   MTPAnalog[2].VExt := 10.0;
   MTPAnalog[0].VOp := 25.0;
   MTPAnalog[1].VOp := 1000.0;
   MTPAnalog[2].VOp := 10.0;
   MTPAnalog[0].VInt := 25.0;
   MTPAnalog[1].VInt := 1000.0;
   MTPAnalog[2].VInt := 10.0;
   MTPAnalog[0].VReq := 25.0;
   MTPAnalog[1].VReq := 1000.0;
   MTPAnalog[2].VReq := 10.0;
   MTPAnalog[0].VOut := 25.0;
   MTPAnalog[1].VOut := 1000.0;
   MTPAnalog[2].VOut := 10.0;
   MTPAnalog[0].VSclMin := 0.0;
   MTPAnalog[1].VSclMin := 100.0;
   MTPAnalog[2].VSclMin := 0.0;
   MTPAnalog[0].VSclMax := 32.0;
   MTPAnalog[1].VSclMax := 3000.0;
   MTPAnalog[2].VSclMax := 300.0;
   MTPAnalog[0].VUnit := 1600;
   MTPAnalog[1].VUnit := 1038;
   MTPAnalog[2].VUnit := 1054;
   MTPAnalog[0].VMin := 0.0;
   MTPAnalog[1].VMin := 100.0;
   MTPAnalog[2].VMin := 5.0;
   MTPAnalog[0].VMax := 32.0;
   MTPAnalog[1].VMax := 3000.0;
   MTPAnalog[2].VMax := 300.0;
END_DATA_BLOCK

DATA_BLOCK "ProcessValues_DB"   // DB34
AUTHOR : Siemens AG
FAMILY : ServiceControl
VERSION : 1.0
// stored: InstanceOfName ProcessValues, InstanceOfType FB
"ProcessValues"
BEGIN
   MTPAnalogIn[0].V := 1500.0;
   MTPAnalogIn[0].SclMinCur := 0.0;
   MTPAnalogIn[0].SclMaxCur := 3000.0;
   MTPAnalogIn[0].UnitCur := 1038;
   MTPAnalogIn[0].SclMinExt := 0.0;
   MTPAnalogIn[0].SclMaxExt := 3000.0;
   MTPAnalogIn[0].UnitExt := 1038;
   MTPBinaryIn[0].V := True;
   MTPBinaryIn[0].VState0 := 'Valve next PEA c';
   MTPBinaryIn[0].VState1 := 'Valve next PEA o';
   MTPAnalogOut[0..1].V := 0.0;
   MTPAnalogOut[0..1].VSclMin := 0.0;
   MTPAnalogOut[0..1].VSclMax := 32.0;
   MTPAnalogOut[0].VUnit := 1351;
   MTPAnalogOut[1].VUnit := 1322;
END_DATA_BLOCK

DATA_BLOCK "ReportValues_DB"   // DB35
AUTHOR : Siemens AG
FAMILY : ServiceControl
VERSION : 1.0
// stored: InstanceOfName ReportValues, InstanceOfType FB
"ReportValues"
BEGIN
   MTPAnalog[0..1].V := 0.0;
   MTPAnalog[0..1].VSclMin := 0.0;
   MTPAnalog[0].VSclMax := 32.0;
   MTPAnalog[1].VSclMax := 100000.0;
   MTPAnalog[0].VUnit := 1351;
   MTPAnalog[1].VUnit := 1038;
END_DATA_BLOCK

DATA_BLOCK "ServiceCommandLogicDB"   // DB11
// stored: InstanceOfName Service_Command_Logic, InstanceOfType FB
"Service_Command_Logic"
BEGIN
END_DATA_BLOCK

DATA_BLOCK "Service_Interaction_FB_DB"   // DB57
// stored: InstanceOfName Service_Interaction_FB, InstanceOfType FB
"Service_Interaction_FB"
BEGIN
END_DATA_BLOCK

DATA_BLOCK "FIC100_Type"   // DB13
// stored: InstanceOfName MTPPIDCtrl_Type1, InstanceOfType FB
"MTPPIDCtrl_Type1"
BEGIN
   AnIn_IDB.Scale.High := 32.0;
   PIDConL_IDB.NegGain.Value := true;
   PIDConL_IDB.Gain.Value := 1.5;
   PIDConL_IDB.TI.Value := 2.0;
   PIDConL_IDB.SP_InHiLim := 32.0;
   PIDConL_IDB.PV_WL_En := false;
   PIDConL_IDB.PV_AL_En := false;
   PIDConL_IDB.RbkWH_En := false;
   PIDConL_IDB.RbkWL_En := false;
   MTPPIDCtrl_IDB.MTP_PIDCtrl.P := 1.5;
   MTPPIDCtrl_IDB.MTP_PIDCtrl.Ti := 2.0;
END_DATA_BLOCK

DATA_BLOCK "FIT100_Type"   // DB2
// stored: InstanceOfName MTPAnaMon_Type1, InstanceOfType FB
"MTPAnaMon_Type1"
BEGIN
   AnIn_IDB.Scale.High := 32.0;
   MonAnL_IDB.PV_AH_Lim := 40.0;
   MonAnL_IDB.PV_WH_Lim := 39.0;
   MonAnL_IDB.PV_TH_Lim := 38.0;
   MonAnL_IDB.PV_TL_Lim := 1.5;
   MonAnL_IDB.PV_WL_Lim := 1.0;
   MonAnL_IDB.PV_AL_Lim := 0.5;
   MonAnL_IDB.PV_AH_En := false;
   MonAnL_IDB.PV_WH_En := false;
   MonAnL_IDB.PV_WL_En := false;
   MonAnL_IDB.PV_AL_En := false;
   MonAnL_IDB.GradHUpEn := false;
   MonAnL_IDB.GradHDnEn := false;
END_DATA_BLOCK

DATA_BLOCK "FIT100Liter_Type"   // DB1
// stored: InstanceOfName MTPAnaMon_Type1, InstanceOfType FB
"MTPAnaMon_Type1"
BEGIN
   AnIn_IDB.Scale.High := 3600.0;
   MonAnL_IDB.PV_AH_En := false;
   MonAnL_IDB.PV_WH_En := false;
   MonAnL_IDB.PV_WL_En := false;
   MonAnL_IDB.PV_AL_En := false;
   MonAnL_IDB.GradHUpEn := false;
   MonAnL_IDB.GradHDnEn := false;
END_DATA_BLOCK

DATA_BLOCK "LAH100_Type"   // DB19
// stored: InstanceOfName MTPBinMon_Type1, InstanceOfType FB
"MTPBinMon_Type1"
BEGIN
END_DATA_BLOCK

DATA_BLOCK "LAL100_Type"   // DB15
// stored: InstanceOfName MTPBinMon_Type1, InstanceOfType FB
"MTPBinMon_Type1"
BEGIN
END_DATA_BLOCK

DATA_BLOCK "LIT100_Type"   // DB12
// stored: InstanceOfName MTPAnaMon_Type1, InstanceOfType FB
"MTPAnaMon_Type1"
BEGIN
   AnIn_IDB.Scale.High := 3000.0;
   MonAnL_IDB.PV_AH_Lim := 2900.0;
   MonAnL_IDB.PV_WH_Lim := 2800.0;
   MonAnL_IDB.PV_TH_Lim := 2700.0;
   MonAnL_IDB.PV_TL_Lim := 150.0;
   MonAnL_IDB.PV_WL_Lim := 90.0;
   MonAnL_IDB.PV_AL_Lim := 30.0;
   MonAnL_IDB.PV_TH_En := true;
   MonAnL_IDB.PV_TL_En := true;
   MonAnL_IDB.GradHUpEn := false;
   MonAnL_IDB.GradHDnEn := false;
END_DATA_BLOCK

DATA_BLOCK "P100_Type"   // DB3
// stored: InstanceOfName MTPMonBinDrv_Type1, InstanceOfType FB
"MTPMonBinDrv_Type1"
BEGIN
   Intlk04_IDB.DataHMI.In01_Text := '';
   Intlk04_IDB.DataHMI.BypIn01 := FALSE;
   Intlk04_IDB.DataHMI.AV01 := 0.0;
   Intlk04_IDB.DataHMI.AV01_Unit := 0;
   Intlk04_IDB.DataHMI.In02_Text := '';
   Intlk04_IDB.DataHMI.BypIn02 := FALSE;
   Intlk04_IDB.DataHMI.AV02 := 0.0;
   Intlk04_IDB.DataHMI.AV02_Unit := 0;
   Intlk04_IDB.DataHMI.In03_Text := '';
   Intlk04_IDB.DataHMI.BypIn03 := FALSE;
   Intlk04_IDB.DataHMI.AV03 := 0.0;
   Intlk04_IDB.DataHMI.AV03_Unit := 0;
   Intlk04_IDB.DataHMI.In04_Text := '';
   Intlk04_IDB.DataHMI.BypIn04 := FALSE;
   Intlk04_IDB.DataHMI.AV04 := 0.0;
   Intlk04_IDB.DataHMI.AV04_Unit := 0;
   Intlk04_IDB.DataHMI.RstOp := FALSE;
   Intlk04_IDB.DataHMI.RstBypOp := FALSE;
   Intlk04_IDB.DataHMI.OS_PermOut := 16#FFFF_FFFF;
   Intlk04_IDB.DataHMI.OS_PermLog := 16#FFF0_FFF9;
   Intlk04_IDB.DataHMI.OpSt_Out := 16#0000_0000;
   Intlk04_IDB.DataHMI.ST_Worst := 16#80;
   Intlk04_IDB.DataHMI.Status1 := 16#0000_0202;
   Intlk04_IDB.DataHMI.Status2 := 16#0000_000E;
   Intlk04_IDB.DataHMI.Status3 := 16#0000_0000;
   Intlk04_IDB.DataHMI.Status4 := 16#0000_000E;
   Intlk04_IDB.DataHMI.Status5 := 16#0000_0000;
   Intlk04_IDB.DataHMI.Status6 := 16#0000_0000;
   Intlk04_IDB.DataHMI.Status7 := 16#0000_000F;
   Intlk04_IDB.DataHMI.Status8 := 16#0000_0000;
   MotL_IDB.Monitor := TRUE;
   MotL_IDB.MonTiStatic := 10.0;
   MotL_IDB.MonTiDynamic := 10.0;
   MotL_IDB.MonTiDyStop := 3.0;
   MotL_IDB.SimOn := FALSE;
   MotL_IDB.DataHMI.StartMan := FALSE;
   MotL_IDB.DataHMI.StopMan := FALSE;
   MotL_IDB.DataHMI.AutModOp := FALSE;
   MotL_IDB.DataHMI.ManModOp := FALSE;
   MotL_IDB.DataHMI.LocalOp := FALSE;
   MotL_IDB.DataHMI.OosOp := FALSE;
   MotL_IDB.DataHMI.LocalLi := FALSE;
   MotL_IDB.DataHMI.StartLocal := FALSE;
   MotL_IDB.DataHMI.StopLocal := FALSE;
   MotL_IDB.DataHMI.Monitor := TRUE;
   MotL_IDB.DataHMI.MonTiStatic := 10.0;
   MotL_IDB.DataHMI.MonTiDynamic := 10.0;
   MotL_IDB.DataHMI.MonTiDyStop := 3.0;
   MotL_IDB.DataHMI.RapidStp := FALSE;
   MotL_IDB.DataHMI.RstOp := FALSE;
   MotL_IDB.DataHMI.Permit_ST := 16#FF;
   MotL_IDB.DataHMI.Intlock_ST := 16#80;
   MotL_IDB.DataHMI.Protect_ST := 16#FF;
   MotL_IDB.DataHMI.CurrMon := 0;
   MotL_IDB.DataHMI.FbkRunOut := FALSE;
   MotL_IDB.DataHMI.OS_PermOut := 16#FFFF_FFFF;
   MotL_IDB.DataHMI.OS_PermLog := 16#7BFF_FF49;
   MotL_IDB.DataHMI.OpSt_Out := 16#0000_0000;
   MotL_IDB.DataHMI.ST_Worst := 16#80;
   MotL_IDB.DataHMI.Status1 := 16#1081_0280;
   MotL_IDB.DataHMI.Status2 := 16#4010_0000;
   MotL_IDB.DataHMI.Status3 := 16#0200_8000;
   MotL_IDB.DataHMI.Status4 := 16#0000_0400;
   MotL_IDB.DataHMI.AlarmState := 16#0000;
   MotL_IDB.Start.Value := FALSE;
   MotL_IDB.Start.InternalUseBit1 := FALSE;
   MotL_IDB.Start.InternalUseBit2 := FALSE;
   MotL_IDB.Start.InternalUseBit3 := FALSE;
   MotL_IDB.Start.InternalUseBit4 := FALSE;
   MotL_IDB.Start.InternalUseBit5 := FALSE;
   MotL_IDB.Start.InternalUseBit6 := FALSE;
   MotL_IDB.Start.InternalUseBit7 := FALSE;
   MotL_IDB.Start.ST := 16#80;
   MotL_IDB.LocalAct.Value := FALSE;
   MotL_IDB.LocalAct.InternalUseBit1 := FALSE;
   MotL_IDB.LocalAct.InternalUseBit2 := FALSE;
   MotL_IDB.LocalAct.InternalUseBit3 := FALSE;
   MotL_IDB.LocalAct.InternalUseBit4 := FALSE;
   MotL_IDB.LocalAct.InternalUseBit5 := FALSE;
   MotL_IDB.LocalAct.InternalUseBit6 := FALSE;
   MotL_IDB.LocalAct.InternalUseBit7 := FALSE;
   MotL_IDB.LocalAct.ST := 16#80;
   MotL_IDB.AutAct.Value := FALSE;
   MotL_IDB.AutAct.InternalUseBit1 := FALSE;
   MotL_IDB.AutAct.InternalUseBit2 := FALSE;
   MotL_IDB.AutAct.InternalUseBit3 := FALSE;
   MotL_IDB.AutAct.InternalUseBit4 := FALSE;
   MotL_IDB.AutAct.InternalUseBit5 := FALSE;
   MotL_IDB.AutAct.InternalUseBit6 := FALSE;
   MotL_IDB.AutAct.InternalUseBit7 := FALSE;
   MotL_IDB.AutAct.ST := 16#80;
   MotL_IDB.ManAct.Value := TRUE;
   MotL_IDB.ManAct.InternalUseBit1 := FALSE;
   MotL_IDB.ManAct.InternalUseBit2 := FALSE;
   MotL_IDB.ManAct.InternalUseBit3 := FALSE;
   MotL_IDB.ManAct.InternalUseBit4 := FALSE;
   MotL_IDB.ManAct.InternalUseBit5 := FALSE;
   MotL_IDB.ManAct.InternalUseBit6 := FALSE;
   MotL_IDB.ManAct.InternalUseBit7 := FALSE;
   MotL_IDB.ManAct.ST := 16#80;
   MotL_IDB.OosAct.Value := FALSE;
   MotL_IDB.OosAct.InternalUseBit1 := FALSE;
   MotL_IDB.OosAct.InternalUseBit2 := FALSE;
   MotL_IDB.OosAct.InternalUseBit3 := FALSE;
   MotL_IDB.OosAct.InternalUseBit4 := FALSE;
   MotL_IDB.OosAct.InternalUseBit5 := FALSE;
   MotL_IDB.OosAct.InternalUseBit6 := FALSE;
   MotL_IDB.OosAct.InternalUseBit7 := FALSE;
   MotL_IDB.OosAct.ST := 16#80;
   MotL_IDB.Run.Value := FALSE;
   MotL_IDB.Run.InternalUseBit1 := FALSE;
   MotL_IDB.Run.InternalUseBit2 := FALSE;
   MotL_IDB.Run.InternalUseBit3 := FALSE;
   MotL_IDB.Run.InternalUseBit4 := FALSE;
   MotL_IDB.Run.InternalUseBit5 := FALSE;
   MotL_IDB.Run.InternalUseBit6 := FALSE;
   MotL_IDB.Run.InternalUseBit7 := FALSE;
   MotL_IDB.Run.ST := 16#80;
   MotL_IDB.Stop.Value := TRUE;
   MotL_IDB.Stop.InternalUseBit1 := FALSE;
   MotL_IDB.Stop.InternalUseBit2 := FALSE;
   MotL_IDB.Stop.InternalUseBit3 := FALSE;
   MotL_IDB.Stop.InternalUseBit4 := FALSE;
   MotL_IDB.Stop.InternalUseBit5 := FALSE;
   MotL_IDB.Stop.InternalUseBit6 := FALSE;
   MotL_IDB.Stop.InternalUseBit7 := FALSE;
   MotL_IDB.Stop.ST := 16#80;
   MotL_IDB.SrMonTime := 10.0;
   MotL_IDB.SxFirstStart := FALSE;
   MotL_IDB.SxCmdStart := FALSE;
   MotL_IDB.SxLastMode := FALSE;
END_DATA_BLOCK

DATA_BLOCK "P101_Type"   // DB20
// stored: InstanceOfName MTPMonBinDrv_Type1, InstanceOfType FB
"MTPMonBinDrv_Type1"
BEGIN
END_DATA_BLOCK

DATA_BLOCK "CalcDoseDB"   // DB6
// stored: InstanceOfName CalcDose, InstanceOfType FB
"CalcDose"
BEGIN
END_DATA_BLOCK

DATA_BLOCK "SimLIT100"   // DB30
// stored: InstanceOfName Level, InstanceOfType FB
"Level"
BEGIN
END_DATA_BLOCK

DATA_BLOCK "V100PT1"   // DB10
// stored: InstanceOfName PT1, InstanceOfType FB
"PT1"
BEGIN
END_DATA_BLOCK

DATA_BLOCK "Volumeflow_DB"   // DB43
// stored: InstanceOfName Volumeflow, InstanceOfType FB
"Volumeflow"
BEGIN
END_DATA_BLOCK

DATA_BLOCK "V100_Type"   // DB61
// stored: InstanceOfName MTPMonAnaVlv_Type1, InstanceOfType FB
"MTPMonAnaVlv_Type1"
BEGIN
   VlvAnL_IDB.RbkHyst := 0.5;
   VlvAnL_IDB.RbkWL_En := TRUE;
   VlvAnL_IDB.RbkWL_MsgEn := false;
   VlvAnL_IDB.NoFbkOpen := TRUE;
   VlvAnL_IDB.NoFbkClose := TRUE;
   VlvAnL_IDB.MonTiStatic := 10.0;
   VlvAnL_IDB.MonTiDynamic := 10.0;
END_DATA_BLOCK
